// TwinCAT 3 PLC project TcProjectBase
// Title: ATI_KOSTAL_AF2024_AUDI2026_TcProjectBase
// Company: ATI
// Author: Ivana Mishevska
// ProjectVersion: 1.1.0.2
// Description: New library for Festo CMT Drive
// ProgramVersion: 3.1.4024.0
// libraries:
//   KOSTAL.AF2024.Core.FileLogger, * (KOSTAL GmbH & Co.KG)
//   KOSTAL.AF2024.Core.GetSystemTime, * (KOSTAL GmbH & Co.KG)
//   KOSTAL.AF2024.Core.MainControl, * (KOSTAL GmbH & Co.KG)
//   KOSTAL.AF2024.Core.Process, * (KOSTAL GmbH & Co.KG)
//   KOSTAL.AF2024.Core.Settings, * (KOSTAL GmbH & Co.KG)
//   KOSTAL.AF2024.Core.Station, * (KOSTAL GmbH & Co.KG)
//   KOSTAL.AF2024.Core.StringTools, * (KOSTAL GmbH & Co.KG)
//   KOSTAL.AF2024.Core.Text, * (KOSTAL GmbH & Co.KG)
//   KOSTAL.AF2024.Drivers.Actuation.Axis.Festo.CMMT_AS, * (KOSTAL GmbH & Co.KG)
//   KOSTAL.AF2024.Drivers.Actuation.Cylinder, * (KOSTAL GmbH & Co.KG)
//   KOSTAL.AF2024.Drivers.Camera.Cognex_InSight, * (KOSTAL GmbH & Co.KG)
//   KOSTAL.AF2024.Drivers.Camera.I_Camera, * (KOSTAL GmbH & Co.KG)
//   KOSTAL.AF2024.Drivers.Camera.Keyence_IV, * (KOSTAL GmbH & Co.KG)
//   KOSTAL.AF2024.Drivers.Scanner.Cognex.DM260, * (KOSTAL GmbH & Co.KG)
//   KOSTAL.AF2024.Drivers.Scanner.IScanner, * (KOSTAL GmbH & Co.KG)
//   KOSTAL.AF2024.Drivers.Scanner.Keyence_SR, * (KOSTAL GmbH & Co.KG)
//   KOSTAL.AF2024.HMI.I_Hmi, * (KOSTAL GmbH & Co.KG)
//   KOSTAL.AF2024.HMI.WinHMI, * (KOSTAL GmbH & Co.KG)
//   KOSTAL.AF2024.Misc.Counter, * (KOSTAL GmbH & Co.KG)
//   KOSTAL.AF2024.Templates.TextMaster, * (KOSTAL GmbH & Co.KG)
//   KOSTAL.TC3.Device.Axis.FESTO.CMMT_AS.ETC, * (KOSTAL GmbH & Co.KG)
//   Tc2_Standard, * (Beckhoff Automation GmbH)
//   Tc2_System, * (Beckhoff Automation GmbH)
//   Tc2_TcpIp, * (Beckhoff Automation GmbH)
//   Tc2_Utilities, * (Beckhoff Automation GmbH)
//   Tc3_Module, * (Beckhoff Automation GmbH)
//   TcCamera, * (TcNexa)
//   TcCameraKeyenceIX, * (TcNexa)
//   TcProcess, * (TcNexa)
// project tree:
//   00_MainControl_Cell/ FB_MainControlCell.TcPOU, T_E_text_MainControl.TcPOU
//   01_Interface/ I_CustomStationInterface.TcIO
//   02_ControlledStations/ FB_StationBase.TcPOU, FB_StationBaseWithAutomaticSlider.TcPOU, FB_StationBaseWithSlider.TcPOU
//   03_FreeStations/01_Safety/DUTs/ T_E_text_Safety.TcPOU
//   03_FreeStations/01_Safety/ FB_Safety_ST80.TcPOU, FB_SafetyBase.TcPOU, FB_Safety_STAudi.TcPOU, FB_Safety_ST50.TcPOU
//   03_FreeStations/01_Safety/ITFs/ I_Safety.TcIO
//   03_FreeStations/02_Parameters/DUTs/ E_Parameters.TcDUT
//   03_FreeStations/02_Parameters/ FB_ParameterHandler.TcPOU
//   03_FreeStations/02_Parameters/ITFs/ I_Parameters_MainControl.TcIO
//   03_FreeStations/03_TextMaster/DUTs/ T_E_text_Common.TcPOU
//   03_FreeStations/03_TextMaster/ FB_TextMaster.TcPOU
//   03_FreeStations/04_EtherCAT Monitoring/DUTs/ T_E_text_EtherCAT.TcPOU
//   03_FreeStations/04_EtherCAT Monitoring/ FB_EtherCAT_Base.TcPOU
//   03_FreeStations/04_EtherCAT Monitoring/ITFs/ I_EtherCAT.TcIO
//   03_FreeStations/05_Fuse Monitorning/DUTs/ T_E_text_Fuse.TcPOU
//   03_FreeStations/05_Fuse Monitorning/ FB_FuseMonitoringBase.TcPOU
//   03_FreeStations/05_Fuse Monitorning/ITFs/ I_Fuse.TcIO
//   04_ComponentSource/ FB_CounterHandler.TcPOU
//   / GVL_Base_FilesAndFolders.TcGVL, MAIN.TcPOU
//   Version/ Global_Version.TcGVL
// real-time tasks:
//   TASK PlcTask: cycle T#10ms, priority 20, ADS port 350
//   TASK PlcTask1: cycle T#10ms, priority 21, ADS port 351

// ---- 03_FreeStations/02_Parameters/DUTs/E_Parameters.TcDUT
{attribute 'qualified_only'}
{attribute 'strict'}
TYPE E_Parameters :
(
	isLoggerEnabled 				:= 1,
	cylinderTimeout					:= 2,
//	airPressureMin					:= 3,
//	airPressureMax					:= 4,
	numberOfRetries					:= 5
	
);
END_TYPE

// ---- GVL_Base_FilesAndFolders.TcGVL
{attribute 'qualified_only'}
VAR_GLOBAL CONSTANT
	PATH_TEXT_MAIN_CONTROL		: KOSTAL_AF2024_Core_Settings.T_MaxString_UTF8:= 'D:\PLC\Text\MainControl\';
	PATH_TEXT_SAFETY			: KOSTAL_AF2024_Core_Settings.T_MaxString_UTF8:= 'D:\PLC\Text\Safety\';
	PATH_TEXT_ETHERCAT			: KOSTAL_AF2024_Core_Settings.T_MaxString_UTF8:= 'D:\PLC\Text\EtherCAT\';
	PATH_TEXT_FUSE				: KOSTAL_AF2024_Core_Settings.T_MaxString_UTF8:= 'D:\PLC\Text\FuseMonitoring\';
	PATH_PARAMETER_VALUES		: KOSTAL_AF2024_Core_Settings.T_MaxString_UTF8:= 'D:\PLC\Data\parameterValues.json';
	PATH_TEXT_COMMON			: KOSTAL_AF2024_Core_Settings.T_MaxString_UTF8:= 'D:\PLC\Text\Common\';
	PATH_TEXT_MASTER			: KOSTAL_AF2024_Core_Settings.T_MaxString_UTF8:= 'D:\PLC\Text\TextMaster\';
	PATH_TEXT_ARTICLE			: KOSTAL_AF2024_Core_Settings.T_MaxString_UTF8:= 'D:\PLC\Text\Article\';
	PATH_ARTICLES				: KOSTAL_AF2024_Core_Settings.T_MaxString_UTF8:= 'D:\PLC\Article';
	PATH_RESET_COUNTER			: KOSTAL_AF2024_Core_Settings.T_MaxString_UTF8:= 'D:\PLC\Counter\ResettableCounter.json';
	PATH_TOTAL_COUNTER			: KOSTAL_AF2024_Core_Settings.T_MaxString_UTF8:= 'D:\PLC\Counter\TotalCounter.json';
	PATH_LOGGER_PROCESS			: KOSTAL_AF2024_Core_Settings.T_MaxString_UTF8:= 'D:\Log\Process\';
	PATH_LOGGER_SAFETY			: KOSTAL_AF2024_Core_Settings.T_MaxString_UTF8:= 'D:\Log\Safety\';
	PATH_LOGGER_ETHERCAT		: KOSTAL_AF2024_Core_Settings.T_MaxString_UTF8:= 'D:\Log\EtherCAT Diagnostics\';
	PATH_LOGGER_FUSE			: KOSTAL_AF2024_Core_Settings.T_MaxString_UTF8:= 'D:\Log\Fuse Diagnostics\';
	




//	PATH_TEXT_MAIN_CONTROL		: KOSTAL_AF2024_Core_Settings.T_MaxString_UTF8:= 'C:\Users\ATI\Desktop\ST80\PLC\Text\MainControl\';//'D:\PLC\Text\MainControl\';//
//	PATH_TEXT_SAFETY			: KOSTAL_AF2024_Core_Settings.T_MaxString_UTF8:= 'C:\Users\ATI\Desktop\ST80\PLC\Text\Safety\';//'D:\PLC\Text\Safety\';//'
//	PATH_TEXT_ETHERCAT			: KOSTAL_AF2024_Core_Settings.T_MaxString_UTF8:= 'C:\Users\ATI\Desktop\ST80\PLC\Text\EtherCAT\';//'D:\PLC\Text\EtherCAT\';//
//	PATH_TEXT_FUSE				: KOSTAL_AF2024_Core_Settings.T_MaxString_UTF8:= 'C:\Users\ATI\Desktop\ST80\PLC\Text\FuseMonitoring\';//'D:\PLC\Text\FuseMonitoring\';//
//	PATH_PARAMETER_VALUES		: KOSTAL_AF2024_Core_Settings.T_MaxString_UTF8:= 'C:\Users\ATI\Desktop\ST80\PLC\Data\parameterValues.json';//'D:\PLC\Data\parameterValues.json';//
//	PATH_TEXT_COMMON			: KOSTAL_AF2024_Core_Settings.T_MaxString_UTF8:= 'C:\Users\ATI\Desktop\ST80\PLC\Text\Common\';//'D:\PLC\Text\Common\';//
//	PATH_TEXT_MASTER			: KOSTAL_AF2024_Core_Settings.T_MaxString_UTF8:= 'C:\Users\ATI\Desktop\ST80\PLC\Text\TextMaster\';//'D:\PLC\Text\TextMaster\';//
//	PATH_TEXT_ARTICLE			: KOSTAL_AF2024_Core_Settings.T_MaxString_UTF8:= 'C:\Users\ATI\Desktop\ST80\PLC\Text\Article\';//'D:\PLC\Text\Article\';//
//	PATH_ARTICLES				: KOSTAL_AF2024_Core_Settings.T_MaxString_UTF8:= 'C:\Users\ATI\Desktop\ST80\PLC\Article';//'D:\PLC\Article';//
//	PATH_RESET_COUNTER			: KOSTAL_AF2024_Core_Settings.T_MaxString_UTF8:= 'C:\Users\ATI\Desktop\ST80\PLC\Counter\ResettableCounter.json';//
//	PATH_TOTAL_COUNTER			: KOSTAL_AF2024_Core_Settings.T_MaxString_UTF8:= 'D:\PLC\Counter\TotalCounter.json';//'C:\Users\ATI\Desktop\ST80\PLC\Counter\TotalCounter.json';//'D:\PLC\Counter\ResettableCounter.json';//
//	PATH_LOGGER_PROCESS			: KOSTAL_AF2024_Core_Settings.T_MaxString_UTF8:= 'C:\Users\ATI\Desktop\ST80\Log\Process\';//'D:\Log\Process\';//
//	PATH_LOGGER_SAFETY			: KOSTAL_AF2024_Core_Settings.T_MaxString_UTF8:= 'C:\Users\ATI\Desktop\ST80\Log\Safety\';//'D:\Log\Safety\';//
//	PATH_LOGGER_ETHERCAT		: KOSTAL_AF2024_Core_Settings.T_MaxString_UTF8:= 'C:\Users\ATI\Desktop\ST80\Log\EtherCAT Diagnostics\';//'D:\Log\EtherCAT Diagnostics\';//
//	PATH_LOGGER_FUSE			: KOSTAL_AF2024_Core_Settings.T_MaxString_UTF8:= 'C:\Users\ATI\Desktop\ST80\Log\Fuse Diagnostics\';//'D:\Log\Fuse Diagnostics\';//
	
END_VAR

// ---- Version/Global_Version.TcGVL
{attribute 'TcGenerated'}
{attribute 'no-analysis'}
{attribute 'linkalways'}
// This function has been automatically generated from the project information.
VAR_GLOBAL CONSTANT
	{attribute 'const_non_replaced'}
	stLibVersion_ATI_KOSTAL_AF2024_AUDI2026_TcProjectBase : ST_LibVersion := (iMajor := 1, iMinor := 1, iBuild := 0, iRevision := 2, nFlags := 0, sVersion := '1.1.0.2');
END_VAR

// ---- 01_Interface/I_CustomStationInterface.TcIO
INTERFACE I_CustomStationInterface

PROPERTY pressedAbortButton  : BOOL
GET
END_GET
END_PROPERTY

END_INTERFACE

// ---- 03_FreeStations/01_Safety/ITFs/I_Safety.TcIO
INTERFACE I_Safety

PROPERTY PUBLIC doorLock : BOOL
GET
END_GET
SET
END_SET
END_PROPERTY

PROPERTY inHold : BOOL
GET
END_GET
END_PROPERTY

PROPERTY isDoorSafe : BOOL
GET
END_GET
END_PROPERTY

PROPERTY isDoorUsed : BOOL
GET
END_GET
END_PROPERTY

PROPERTY isSafe : BOOL
GET
END_GET
END_PROPERTY

END_INTERFACE

// ---- 03_FreeStations/02_Parameters/ITFs/I_Parameters_MainControl.TcIO
INTERFACE I_Parameters_MainControl

PROPERTY cylinderSensorTimeout : TIME
GET
END_GET
END_PROPERTY

PROPERTY isLoggerEnabled : BOOL
GET
END_GET
END_PROPERTY

PROPERTY numberOfRetries : INT
GET
END_GET
END_PROPERTY

END_INTERFACE

// ---- 03_FreeStations/04_EtherCAT Monitoring/ITFs/I_EtherCAT.TcIO
INTERFACE I_EtherCAT

PROPERTY inError : BOOL
GET
END_GET
END_PROPERTY

END_INTERFACE

// ---- 03_FreeStations/05_Fuse Monitorning/ITFs/I_Fuse.TcIO
INTERFACE I_Fuse

PROPERTY inError : BOOL
GET
END_GET
END_PROPERTY

END_INTERFACE

// ---- 00_MainControl_Cell/FB_MainControlCell.TcPOU
FUNCTION_BLOCK FB_MainControlCell EXTENDS KOSTAL_AF2024_Core_MainControl.FB_MainControl IMPLEMENTS I_CustomStationInterface 
VAR
(*------------------------------------------------------------------------------------------*)
	(* General *)
	_textPath						: KOSTAL_AF2024_Core_Settings.T_MaxString_UTF8;
	_Text							: KOSTAL_AF2024_Core_Text.FB_Handler_Slave;
	_E_Text							: T_E_text_MainControl;
	_setLogRequest					: BOOL;
	_addressHome					: INT;
	_stepDescription				: WSTRING;
	_articleAutoSelection			: BOOL;
	_timerStationsInHome			: Tc2_Standard.TON;
	_tempText						: WSTRING;
	_onAbortButton					: Tc2_Standard.R_TRIG;
//	_pressedAbortButton				: BOOL; 
(*------------------------------------------------------------------------------------------*)
	(* Interface *)
	_IetherCAT						: I_EtherCAT;
	_IfuseMonitroing				: I_Fuse;
	_ISafety						: I_Safety; 
(*------------------------------------------------------------------------------------------*)	 
	(* Hmi *)
	_Hmi							: KOSTAL_AF2024_HMI_WinHMI.FB_MainControl;
	_Hmi_station					: KOSTAL_AF2024_HMI_WinHMI.FB_Page_Station;
(*------------------------------------------------------------------------------------------*)
	(* Mode *)
	_Message						: KOSTAL_AF2024_Core_Process.T_messageText_3_lines;
	_modeAutomaticRequest			: BOOL:= TRUE;
	_modeManualRequest				: BOOL;
	_dataModeRequest				: BOOL;
(*------------------------------------------------------------------------------------------*)
	(* Links *)
	_Ilogger						: KOSTAL_AF2024_Core_FileLogger.I_Logger;
	_Iparameters					: I_Parameters_MainControl;
(*------------------------------------------------------------------------------------------*)
	(* Inputs *)
//	DI_KeySwitch					AT %I* : BOOL;
	DI_KeySwitchAutomatic			AT %I* : BOOL; //2 
	DI_KeySwitchManual				AT %I* : BOOL; //1 
	DI_CheckPressure_PT1			AT %I* : BOOL;
	DI_AbortButton				 	AT %I* : BOOL;
	(* Outputs *)
	DO_AirSupplyOn					AT %Q* : BOOL;
	DO_ReleMainValve_V1				AT %Q* : BOOL;
	DO_ReleMainValve_V2				AT %Q* : BOOL;
	(* Andon Light *)
	DO_AndonLightGreenLamp			AT %Q* : BOOL;
	DO_AndonLightYellowLamp			AT %Q* : BOOL;
	DO_AndonLightRedLamp			AT %Q* : BOOL;
(*------------------------------------------------------------------------------------------*)
END_VAR

VAR CONSTANT
	_STEP_OFF	: INT:= 0;
END_VAR

METHOD PROTECTED _a0_PowerOff
VAR
	_Participant : KOSTAL_AF2024_Core_Settings.T_MaxString;
END_VAR
IF _Step.toggle THEN
	_Message.clear();
	_Hmi.clear();
	_demand.SetUnique_PowerOff();
//	DO_AirSupplyOn:= FALSE;
	DO_ReleMainValve_V1:= FALSE;
	DO_ReleMainValve_V2:= FALSE;
	_setLogRequest:= TRUE;
	_stepDescription:= "PowerOff";
END_IF

// Log
IF _setLogRequest AND _isLogReady() AND _Text.State.ready AND (_Text.LoadedLanguage <> '') THEN
	IF _Log("===START===") THEN 
		_Log(_Text.GetText(Number:= _E_text.off));	
		_setLogRequest:= FALSE;	
	END_IF
END_IF

// Hmi
_Hmi.Button_OnOff.Visible:= FALSE;

IF NOT _Text.State.ready THEN
	_updateHmiText(
		userMessage		:= _Text.GetText(Number:= _E_Text.textHandlerIsNotReady),
		userAction		:= _Text.State.description,
		isErrorMessage	:= FALSE);
ELSIF NOT _Isafety.isSafe THEN
	_updateHmiText(
		userMessage		:= _Text.GetText(Number:= _E_Text.safetyInError),
		userAction		:= "",
		isErrorMessage	:= FALSE);
ELSIF NOT _all_PowerOff(_Participant) THEN
	_updateHmiText(
		userMessage		:= _Text.GetText(Number:= _E_Text.waitForAllOff),
		userAction		:= _Participant,
		isErrorMessage	:= FALSE);
//ELSIF _isAirPressureOk() THEN
//	_Text.ClearVars();
//	_Text.AddVar(Text:= "-1AZ1");
//	_Text.AddVar(Text:= _Text.GetText(Number:= _E_Text.active));
//	_updateHmiText(
//		userMessage		:= _Text.GetText(Number:= _E_Text.systemAirPressure_0_is_1),
//		userAction		:= "",
//		isErrorMessage	:= FALSE);
ELSIF NOT _mode.manual THEN
	_updateHmiText(
		userMessage		:= _Text.GetText(Number:= _E_Text.setManualMode),
		userAction		:= "",
		isErrorMessage	:= FALSE);
ELSE
	_Hmi.Button_OnOff.Visible:= _mode.manual AND NOT _condition.isError();
	
	_Text.ClearVars();
	_Text.AddVar(Text:= _Hmi.Button_OnOff.Text);
	_updateHmiText(
		userMessage		:= _Text.GetText(Number:= _E_Text.onWith_0),
		userAction		:= "",
		isErrorMessage	:= FALSE);

	IF _modeManualRequest AND _Hmi.Button_OnOff.Pulse AND NOT _condition.isError() THEN
		_Step.INC();
	END_IF
END_IF
END_METHOD

METHOD PROTECTED _a1_PowerOn
VAR
	_Participant : KOSTAL_AF2024_Core_Settings.T_MaxString;
END_VAR
IF _step.toggle THEN
	_Hmi.clear();
	_Message.clear();
	_demand.SetUnique_PowerOn();
//	DO_AirSupplyOn:= TRUE;
	DO_ReleMainValve_V1:= TRUE;
	DO_ReleMainValve_V2:= TRUE;
	_log(Text:= _Text.GetText(Number:= _E_Text.powerOn));
	_stepDescription:= "PowerOn";
END_IF

_Hmi.Button_OnOff.Text:= _Text.GetText(Number:= _E_Text.waitForPowerOn);
_Hmi.Button_OnOff.Visible:= TRUE;

//IF NOT _isAirPressureOk() THEN
//	_Text.ClearVars();
////	_Text.AddVar(Text:= INT_TO_WSTRING(_Iparameters.airPressureMin));
////	_Text.AddVar(Text:= INT_TO_WSTRING(AI_AirPressure));
////	_Text.AddVar(Text:= INT_TO_WSTRING(_Iparameters.airPressureMax));
//	_updateHmiText(
//		userMessage		:= _Text.GetText(Number:= _E_Text.waitForAirPressure_0_1_2),
//		userAction		:= "",
//		isErrorMessage	:= FALSE);
IF NOT DI_CheckPressure_PT1 THEN 
	_updateHmiText(
		userMessage		:= "Check pressure",//_Text.GetText(Number:= _E_Text.waitForAirPressure_0_1_2),
		userAction		:= "PT1",
		isErrorMessage	:= FALSE);
ELSIF NOT _all_PowerOn(_Participant) THEN
	_updateHmiText(
		userMessage		:= _Text.GetText(Number:= _E_Text.waitForAllOn),
		userAction		:= _Participant,
		isErrorMessage	:= FALSE);
ELSIF NOT _mode.automatic THEN
	_updateHmiText(
		userMessage		:= _Text.GetText(Number:= _E_Text.setAutomaticMode),
		userAction		:= "",
		isErrorMessage	:= FALSE);
ELSE
	_step.INC();
END_IF
END_METHOD

METHOD PROTECTED _a2_OnToHome
VAR
	_Participant : KOSTAL_AF2024_Core_Settings.T_MaxString;
END_VAR
IF _step.toggle THEN
	_Hmi.clear();
	_demand.SetUnique_OnToHome();
	_log(Text:= _Text.GetText(Number:= _E_Text.onToHomeReleased));
	_stepDescription:= "OnToHome";
END_IF

_Hmi.Button_OnOff.Text:= _Text.GetText(Number:= _E_Text.off);
_Hmi.Button_OnOff.Visible:= TRUE;

IF NOT _all_Home(_Participant) THEN
	_updateHmiText(
		userMessage		:= _Text.GetText(Number:= _E_Text.waitFromHome),
		userAction		:= _Participant,
		isErrorMessage	:= FALSE);
ELSE
	_step.INC();
END_IF
END_METHOD

METHOD PROTECTED _a3_Home
VAR
	_Participant: KOSTAL_AF2024_Core_Settings.T_MaxString;
END_VAR
IF _step.toggle THEN
	_addressHome:= _step.actual;
	_Message.clear();
	_Hmi.clear();
	_demand.SetUnique_Home();
	_log(Text:= _Text.GetText(Number:= _E_Text.stop));
	_stepDescription:= "Home";
END_IF

_Hmi.Button_OnOff.Text:= _Text.GetText(Number:= _E_Text.off);
_Hmi.Button_OnOff.Visible:= TRUE;
_Hmi.Button_RunStop.Text:= _Text.GetText(Number:= _E_Text.start);
_Hmi.Button_RunStop.Visible:= FALSE;

IF NOT _all_Home(_Participant) THEN
	_updateHmiText(
		userMessage		:= _Text.GetText(Number:= _E_Text.participantNotReady),
		userAction		:= _Participant,
		isErrorMessage	:= FALSE);
ELSIF _Hmi.Button_RunStop.Pulse OR NOT _enableStopMode THEN
	_Hmi.Button_RunStop.Visible:= FALSE;
	_step.INC();
ELSE
	_Hmi.Button_RunStop.Visible:= TRUE;
	_updateHmiText(
		userMessage		:= _Text.GetText(Number:= _E_Text.stop),
		userAction		:= _Text.GetText(Number:= _E_Text.readyToStart),
		isErrorMessage	:= FALSE);
END_IF
END_METHOD

METHOD PROTECTED _a4_Run
VAR_INPUT
END_VAR
IF _step.toggle THEN
	_Hmi.clear();
	_demand.SetUnique_Run();
	_log(Text:= _Text.GetText(Number:= _E_Text.busy));
	_stepDescription:= "Run";
END_IF

_Hmi.Button_OnOff.Text:= _Text.GetText(Number:= _E_Text.off);
_Hmi.Button_OnOff.Visible:= TRUE;
_Hmi.Button_RunStop.Text:= _Text.GetText(Number:= _E_Text.stop);
_Hmi.Button_RunStop.Visible:= _enableStopMode;

IF _Hmi.Button_RunStop.Pulse AND _enableStopMode THEN
	_step.INC();
//ELSIF NOT _isAirPressureOk() THEN
//	_updateHmiText(
//		userMessage		:= "Air pressure out of limits",
//		userAction		:= "",
//		isErrorMessage	:= TRUE);
//	_step.init();	
//ELSIF (_IetherCAT <> 0) AND_THEN _IetherCAT.inError THEN
//	_updateHmiText(
//		userMessage		:= "EtherCAT in fault",
//		userAction		:= "",
//		isErrorMessage	:= TRUE);
//	_step.init();	
//ELSIF (_IfuseMonitroing <> 0) AND_THEN _IfuseMonitroing.inError THEN
//	_updateHmiText(
//		userMessage		:= "Fuse in fault",
//		userAction		:= "",
//		isErrorMessage	:= TRUE);
//	_step.init();	
ELSE
	_tempText:= "";
//	IF (_IArticle <> 0) THEN
//		IF _IArticle.LoadedArticle.isVariantTypeGen6x THEN
//			_tempText:= "Selected article: Gen6x";
//		ELSIF _IArticle.LoadedArticle.isProductTypeGen6 THEN
//			_tempText:= "Selected article: Gen6";
//		ELSIF _IArticle.LoadedArticle.isProductTypeGen7 THEN
//			_tempText:= "Selected article: Gen7";
//		ELSIF _IArticle.LoadedArticle.isProductTypeVan THEN
//			_tempText:= "Selected article: Van";
//		END_IF
//	END_IF

	_updateHmiText(
		userMessage		:= _Text.GetText(Number:= _E_Text.run),
		userAction		:= _tempText,
		isErrorMessage	:= FALSE);
END_IF
END_METHOD

METHOD PROTECTED _a5_RunToHome
VAR
	_Participant: KOSTAL_AF2024_Core_Settings.T_MaxString;
END_VAR
IF _step.toggle THEN
	_Message.clear();
	_Hmi.clear();
	_demand.SetUnique_RunToHome();
	_log(Text:= _Text.GetText(Number:= _E_Text.lastCycle));
	_stepDescription:= "RunToHome";
END_IF

_Hmi.Button_OnOff.Text:= _Text.GetText(Number:= _E_Text.off);
_Hmi.Button_OnOff.Visible:= TRUE;
_Hmi.Button_RunStop.Text:= _Text.GetText(Number:= _E_Text.start);
_Hmi.Button_RunStop.Visible:= TRUE;

IF _Hmi.Button_RunStop.Pulse OR NOT _enableStopMode THEN
	_step.DEC();
ELSIF _all_Home(_Participant) THEN
	_step.set(request:= _addressHome);
ELSE
	_updateHmiText(
		userMessage		:= _Text.GetText(Number:= _E_Text.participantNotReady),
		userAction		:= _Participant,
		isErrorMessage	:= FALSE);
END_IF
END_METHOD

METHOD PROTECTED _aX_Fail
VAR_INPUT
END_VAR
_demand.clear();

_Message.clear();
_Text.ClearVars();
_Text.AddVar(Text:= INT_TO_WSTRING(_Step.actual));
_Message.line_01:= _Text.GetText(Number:= _E_Text.step_0_doesNotExist);
_condition.setMessage(
	priority:= _condition.PriorityLevel_Error + 1000,
	message:= _Message);
	
IF _Step.toggle THEN
	_Log(Text:= _Message.toString());
END_IF

_Step.init();
END_METHOD

METHOD PROTECTED _checkIfSamePosition : BOOL
VAR_INPUT
	actualPosition 			: LREAL;
	targetPosotion			: LREAL;
END_VAR
IF (actualPosition >= (targetPosotion - 1)) AND (actualPosition <= (targetPosotion + 1)) THEN 
	_checkIfSamePosition:= TRUE;
ELSE 
	_checkIfSamePosition:= FALSE;
END_IF
END_METHOD

METHOD PROTECTED _getIdAsString : KOSTAL_AF2024_Core_Settings.T_MaxString
VAR
	_temp 		: KOSTAL_AF2024_Core_StringTools.FB_Concat;
END_VAR
_temp.Clear();
_temp.addContent(Text:= _ID.name);
_temp.addContent(Text:= "(");
_temp.addContent(Text:= DINT_TO_WSTRING(_ID.key));
_temp.addContent(Text:= ")");
_getIdAsString:= _temp.getResult();
_temp.Clear();
END_METHOD

METHOD PROTECTED _globalError
VAR_INPUT
END_VAR
END_METHOD

METHOD PROTECTED _handleAndonLight
VAR
	_Participant	: KOSTAL_AF2024_Core_Settings.T_MaxString;
END_VAR
IF NOT _Isafety.isSafe THEN
	_timerStationsInHome(IN:= FALSE);
	DO_AndonLightGreenLamp:= FALSE;
	DO_AndonLightYellowLamp:= FALSE;
	DO_AndonLightRedLamp:= TRUE;
ELSIF _mode.manual THEN
	_timerStationsInHome(IN:= FALSE);
	DO_AndonLightGreenLamp:= FALSE;
	DO_AndonLightYellowLamp:= TRUE;
	DO_AndonLightRedLamp:= FALSE;
ELSIF _all_Home(_Participant) THEN
	_timerStationsInHome(IN:= TRUE, PT:= T#1S);
	DO_AndonLightYellowLamp:= FALSE;
	DO_AndonLightRedLamp:= FALSE;
	IF _timerStationsInHome.Q THEN
		_timerStationsInHome(IN:= FALSE);
		DO_AndonLightGreenLamp:= NOT DO_AndonLightGreenLamp;
	END_IF
ELSE
	_timerStationsInHome(IN:= FALSE);
	DO_AndonLightGreenLamp:= TRUE;
	DO_AndonLightYellowLamp:= FALSE;
	DO_AndonLightRedLamp:= FALSE;
END_IF
END_METHOD

METHOD PROTECTED _hmiDefine
VAR
	_Participant: KOSTAL_AF2024_Core_Settings.T_MaxString;
END_VAR
_Hmi.FBmain();
_Hmi_station.FBmain();

// General
_Hmi.Name:= "";
_Hmi.linkMainControl(THIS^);

_Hmi_station.Name:= Tc2_Standard.WCONCAT(
	STR1:= _Text.GetText(Number:= _E_Text.name),
	STR2:= " [");
_Hmi_station.Name:= Tc2_Standard.WCONCAT(
	STR1:= _Hmi_station.Name,
	STR2:= STRING_TO_WSTRING(stLibVersion_ATI_KOSTAL_AF2024_AUDI2026_TcProjectBase.sVersion));
_Hmi_station.Name:= Tc2_Standard.WCONCAT(
	STR1:= _Hmi_station.Name,
	STR2:= "]");

// Mode handling
_mode.manual:= _modeManualRequest;
_mode.automatic:= _modeAutomaticRequest AND NOT _Isafety.inHold;

// Buttons 
_Hmi.Button_Parameters.Visible:= (NOT DI_KeySwitchAutomatic AND NOT DI_KeySwitchManual) AND _dataModeRequest;//_mode.automatic
_Hmi.Button_Article.Visible:= _mode.manual AND _demand.Run; //AND (_Hmi.UserLevel >= KOSTAL_AF2024_HMI_I_Hmi.E_UserLevel.service);
_Hmi.Button_RunStop.Visible:= _enableStopMode;
_Hmi.ManualDeviceControl:= _mode.manual AND _demand.Run AND (_Hmi.UserLevel >= KOSTAL_AF2024_HMI_I_Hmi.E_UserLevel.service);


_Hmi.Button_Door.Visible:= _ISafety.isDoorUsed;
IF _Hmi.Button_Door.Pulse THEN
	_ISafety.doorLock:= NOT _ISafety.doorLock;
END_IF
_Hmi.statusDoor_safe:= _ISafety.isDoorSafe;

_Hmi_station.Button_Escape.Visible:= _condition.isError() AND _modeManualRequest;
_Hmi_station.Button_Escape.Text:= _Text.GetText(Number:= _E_Text.reset);

// Message
_Hmi_station.Text.line_01:= _condition.Message.line_01;
_Hmi_station.Text.line_02:= _condition.Message.line_02;
_Hmi_station.Text.line_03:= _condition.Message.line_03;
_Hmi_station.Status.CopyFrom(IN:= _condition);
END_METHOD

METHOD PROTECTED _isLogReady  : BOOL
VAR_INPUT
END_VAR
IF (_Ilogger = 0) THEN RETURN; END_IF
_isLogReady:= _Ilogger.State.success;
END_METHOD

METHOD PROTECTED _log : BOOL
VAR_INPUT
	Text			  : KOSTAL_AF2024_Core_Settings.T_MaxString;
END_VAR
IF (Text = "") THEN RETURN; END_IF
IF (_Iparameters <> 0) AND_THEN NOT _Iparameters.isLoggerEnabled THEN RETURN; END_IF
IF (_Ilogger = 0) THEN RETURN; END_IF
IF NOT _Ilogger.State.success THEN RETURN; END_IF

_Ilogger.ID:= _getIdAsString();
_Ilogger.name:= _Text.GetText(Number:= _E_Text.name);
_Ilogger.stepNumber:= _Step.actual;

_log:= _Ilogger.addLine(line:= Text);
END_METHOD

METHOD _modeHandler
VAR_INPUT
END_VAR
_mode.automatic:= (_modeAutomaticRequest OR DI_KeySwitchAutomatic) AND NOT _condition.isError() AND NOT _Isafety.inHold AND NOT _dataModeRequest; 
_mode.manual:= _modeManualRequest AND NOT _dataModeRequest;
END_METHOD

METHOD PROTECTED _modeRequest
VAR_INPUT
END_VAR
_Hmi.Button_Auto.Visible:= TRUE;
_Hmi.Button_Manual.Visible:= TRUE;
IF _Hmi.Button_Auto.Pulse OR DI_KeySwitchAutomatic THEN	
	_modeAutomaticRequest:= TRUE;	
	_modeManualRequest:= FALSE;
	_dataModeRequest:= FALSE;
ELSIF _Hmi.Button_Manual.Pulse OR DI_KeySwitchManual THEN	
	_modeAutomaticRequest:= FALSE;	
	_modeManualRequest:= TRUE;
	_dataModeRequest:= FALSE;
ELSIF NOT DI_KeySwitchAutomatic AND NOT DI_KeySwitchManual THEN 
//	_Hmi.Button_Auto.Visible:= TRUE;
//	_Hmi.Button_Manual.Visible:= TRUE;
	_dataModeRequest:= TRUE;
	_modeAutomaticRequest:= FALSE;
	_modeManualRequest:= FALSE;
END_IF
END_METHOD

METHOD PROTECTED _parameterControl : BOOL
VAR_INPUT
END_VAR
_parameterControl:= TRUE;
END_METHOD

METHOD PROTECTED _resetCondition  
VAR_INPUT
END_VAR
IF _condition.isError() THEN
	IF _Hmi_station.Button_Escape.Pulse THEN
		_condition.clear();
	END_IF
ELSE
	_condition.clear();
END_IF
END_METHOD

METHOD PROTECTED _stepHeader
VAR_INPUT
END_VAR
//Switch off in case of off command or safety error
IF _step.actual > _STEP_OFF THEN
	IF _hmi.Button_OnOff.Pulse THEN	
		_step.init();
	ELSIF NOT _Isafety.IsSafe THEN
		_step.init();
	END_IF
END_IF
//Call Step sequence header
_step.Header();
END_METHOD

METHOD PROTECTED _steps
VAR_INPUT
END_VAR
_stepHeader();

CASE _Step.actual OF
	0:	_a0_PowerOff();
	1:	_a1_PowerOn();
	2:	_a2_OnToHome();
	3:	_a3_Home();
	4:	_a4_Run();
	5:	_a5_RunToHome();
ELSE
	_aX_Fail();
END_CASE
END_METHOD

METHOD PROTECTED _textReader : BOOL
VAR_INPUT
END_VAR
_Text.Path:= _textPath;
_Text.FBmain();

IF _Text.State.fail THEN
	_Message.clear();
	_Message.line_01:= "TextHandler";
	_Message.line_02:= _Text.State.description;
	_condition.setMessage(
		priority:= _condition.PriorityLevel_Error,
		message	:= _Message);
ELSIF NOT _Text.Valid THEN
	_Message.clear();
	_Message.line_01:= "TextHandler";
	_Message.line_02:= _Text.State.description;
	_condition.setMessage(
		priority:= _condition.PriorityLevel_MasterMessage + 999,
		message	:= _Message);
END_IF

IF _Text.LoadedLanguage <> '' THEN
	_textReader:= TRUE;
END_IF
END_METHOD

METHOD PROTECTED _updateHmiText
VAR_INPUT
	userMessage		: WSTRING;
	userAction		: WSTRING;
	isErrorMessage	: BOOL;
END_VAR
_message.clear();

_Text.ClearVars();
_Text.AddVar(Text:= INT_TO_WSTRING(_step.actual));
_Text.AddVar(Text:= _stepDescription);
_Text.AddVar(Text:= "0");
_message.line_01:= _Text.GetText(Number:= _E_Text.step_0_actual_1);
_message.line_02:= userMessage;
_message.line_03:= userAction;
IF isErrorMessage AND NOT _condition.isError() THEN
	_log(Text:= _message.toString());
END_IF

IF isErrorMessage THEN
	_condition.setMessage(
		priority:= _condition.PriorityLevel_Error,
		message	:= _message);
ELSIF (userAction <> "") THEN
	_condition.setMessage(
		priority:= _condition.PriorityLevel_Message,
		message	:= _message);
ELSE
	_condition.setMessage(
		priority:= _condition.PriorityLevel_Text,
		message	:= _message);
END_IF
END_METHOD

PROPERTY articleAutoSelection : BOOL
GET
articleAutoSelection:= _articleAutoSelection;
END_GET
SET
_articleAutoSelection:= articleAutoSelection;
END_SET
END_PROPERTY

METHOD FB_init : BOOL
VAR_INPUT
	bInitRetains 		: BOOL; // if TRUE, the retain variables are initialized (warm start / cold start)
	bInCopyCode 		: BOOL;  // if TRUE, the instance afterwards gets moved into the copy code (online change)
	EnableStopMode		: BOOL;
	CommonText			: KOSTAL_AF2024_Core_Text.I_Text;
	textPath			: KOSTAL_AF2024_Core_Settings.T_MaxString_UTF8;
	Parameters			: I_Parameters_MainControl;
	Safety				: I_Safety;
	EtherCAT			: I_EtherCAT;
	Fuse				: I_Fuse;
	Logger				: KOSTAL_AF2024_Core_FileLogger.I_Logger;
//	Article				: I_Article;
END_VAR
THIS^._enableStopMode:= EnableStopMode;
THIS^._Text.linkCommonText(Common:= CommonText);
THIS^._textPath:= textPath;
THIS^._Iparameters:= Parameters;
THIS^._Isafety:= Safety;
THIS^._IetherCAT:= EtherCAT;
THIS^._IfuseMonitroing:= Fuse;
THIS^._Ilogger:= Logger;
END_METHOD

METHOD PUBLIC FBmain 
VAR_INPUT
END_VAR
_modeRequest();

IF NOT _parameterControl() THEN RETURN; END_IF
_hmiDefine();
_resetCondition();
_handleAndonLight();

IF NOT _TextReader() THEN RETURN; END_IF

_globalError();
_modeHandler();
_steps();

_onAbortButton(CLK:= DI_AbortButton);
END_METHOD

PROPERTY language : KOSTAL_AF2024_HMI_I_Hmi.T_LANGUAGENAME
GET
language:= _Hmi.Language;
END_GET
END_PROPERTY

{warning 'add property implementation'}
PROPERTY pressedAbortButton : BOOL
GET
pressedAbortButton:= _onAbortButton.Q;
END_GET
END_PROPERTY

PROPERTY user : KOSTAL_AF2024_HMI_I_Hmi.E_UserLevel
GET
user:= _Hmi.UserLevel;
END_GET
END_PROPERTY

END_FUNCTION_BLOCK

// ---- 00_MainControl_Cell/T_E_text_MainControl.TcPOU
FUNCTION_BLOCK T_E_text_MainControl EXTENDS KOSTAL_AF2024_Core_Text.T_E_Text
VAR
END_VAR

PROPERTY busy : KOSTAL_AF2024_Core_Text.ST_E_Text
GET
busy.Number:= 36;
END_GET
END_PROPERTY

PROPERTY lastCycle : KOSTAL_AF2024_Core_Text.ST_E_Text
GET
lastCycle.Number:= 37;
END_GET
END_PROPERTY

PROPERTY name : KOSTAL_AF2024_Core_Text.ST_E_Text
GET
name.Number:= 2;
END_GET
END_PROPERTY

PROPERTY nextPage : KOSTAL_AF2024_Core_Text.ST_E_Text
GET
nextPage.Number:= 61;
END_GET
END_PROPERTY

PROPERTY off : KOSTAL_AF2024_Core_Text.ST_E_Text
GET
off.Source:= KOSTAL_AF2024_Core_Text.E_Source.Common;
off.Number:= 2;
END_GET
END_PROPERTY

PROPERTY onToHomeReleased : KOSTAL_AF2024_Core_Text.ST_E_Text
GET
onToHomeReleased.Source:= KOSTAL_AF2024_Core_Text.E_Source.Common;
onToHomeReleased.Number:= 42;
END_GET
END_PROPERTY

PROPERTY onWith_0 : KOSTAL_AF2024_Core_Text.ST_E_Text
GET
onWith_0.Source:= KOSTAL_AF2024_Core_Text.E_Source.Common;
onWith_0.Number:= 65;
END_GET
END_PROPERTY

PROPERTY participantNotReady : KOSTAL_AF2024_Core_Text.ST_E_Text
GET
participantNotReady.Number:= 12;
END_GET
END_PROPERTY

PROPERTY powerOn : KOSTAL_AF2024_Core_Text.ST_E_Text
GET
powerOn.Number:= 44;
END_GET
END_PROPERTY

PROPERTY previousPage : KOSTAL_AF2024_Core_Text.ST_E_Text
GET
previousPage.Number:= 60;
END_GET
END_PROPERTY

PROPERTY readyToStart : KOSTAL_AF2024_Core_Text.ST_E_Text
GET
readyToStart.Number:=35;
END_GET
END_PROPERTY

PROPERTY refresh : KOSTAL_AF2024_Core_Text.ST_E_Text
GET
refresh.Number:= 62;
END_GET
END_PROPERTY

PROPERTY reset : KOSTAL_AF2024_Core_Text.ST_E_Text
GET
reset.Source:= Kostal_AF2024_Core_Text.E_Source.Common;
reset.Number:= 7;
END_GET
END_PROPERTY

PROPERTY run : KOSTAL_AF2024_Core_Text.ST_E_Text
GET
run.Number:= 5;
END_GET
END_PROPERTY

PROPERTY safetyInError : KOSTAL_AF2024_Core_Text.ST_E_Text
GET
safetyInError.Number:= 30;
END_GET
END_PROPERTY

PROPERTY setAutomaticMode : KOSTAL_AF2024_Core_Text.ST_E_Text
GET
setAutomaticMode.Number:=41;
END_GET
END_PROPERTY

PROPERTY setManualMode : KOSTAL_AF2024_Core_Text.ST_E_Text
GET
setManualMode.Number:= 40;
END_GET
END_PROPERTY

PROPERTY start : KOSTAL_AF2024_Core_Text.ST_E_Text
GET
start.Source:= KOSTAL_AF2024_Core_Text.E_Source.Common;
start.Number:= 5;
END_GET
END_PROPERTY

PROPERTY step_0_actual_1 : KOSTAL_AF2024_Core_Text.ST_E_Text
GET
step_0_actual_1.Source:= KOSTAL_AF2024_Core_Text.E_Source.Common;
step_0_actual_1.Number:= 11;
END_GET
END_PROPERTY

PROPERTY step_0_doesNotExist : KOSTAL_AF2024_Core_Text.ST_E_Text
GET
step_0_doesNotExist.Source:= KOSTAL_AF2024_Core_Text.E_Source.Common;
step_0_doesNotExist.Number:= 12;
END_GET
END_PROPERTY

PROPERTY stop : KOSTAL_AF2024_Core_Text.ST_E_Text
GET
stop.Source:= KOSTAL_AF2024_Core_Text.E_Source.Common;
stop.Number:= 4;
END_GET
END_PROPERTY

PROPERTY textHandlerIsNotReady : KOSTAL_AF2024_Core_Text.ST_E_Text
GET
textHandlerIsNotReady.Source:= KOSTAL_AF2024_Core_Text.E_Source.Common;
textHandlerIsNotReady.Number:= 20;
END_GET
END_PROPERTY

PROPERTY waitForAirPressure_0_1_2 : KOSTAL_AF2024_Core_Text.ST_E_Text
GET
waitForAirPressure_0_1_2.Number:= 31;
END_GET
END_PROPERTY

PROPERTY waitForAllOff : KOSTAL_AF2024_Core_Text.ST_E_Text
GET
waitForAllOff.Number:= 10;
END_GET
END_PROPERTY

PROPERTY waitForAllOn : KOSTAL_AF2024_Core_Text.ST_E_Text
GET
waitForAllOn.Number:= 11;
END_GET
END_PROPERTY

PROPERTY waitForPowerOn : KOSTAL_AF2024_Core_Text.ST_E_Text
GET
waitForPowerOn.Number:= 13;
END_GET
END_PROPERTY

PROPERTY waitFromHome : KOSTAL_AF2024_Core_Text.ST_E_Text
GET
waitFromHome.Number:= 43;
END_GET
END_PROPERTY

END_FUNCTION_BLOCK

// ---- 02_ControlledStations/FB_StationBase.TcPOU
FUNCTION_BLOCK ABSTRACT FB_StationBase EXTENDS KOSTAL_AF2024_Core_Station.FB_Station_Controlled 
VAR PERSISTENT
	_isCameraMasterDone					: BOOL;
	_lastCameraMasterTime				: DINT;	
END_VAR                         		
VAR                             		
	(* General *)  	            		
	_Hmi_station						: KOSTAL_AF2024_HMI_WinHMI.FB_Page_Station;
	_E_TextCommon						: T_E_text_Common;
	_IgetTime							: KOSTAL_AF2024_Core_GetSystemTime.I_TimeSource;
	_isDevicesInit						: BOOL;
	_cylinderInManualMode				: BOOL;
	_manualModeInterlock				: BOOL;
	_onPowerOff							: Tc2_Standard.R_TRIG;
	_onNagaraSwitch						: Tc2_Standard.R_TRIG;
//	_onAbortButton						: Tc2_Standard.R_TRIG;
	_timerCycleTimer					: Tc2_Standard.TON;
	_addressRestart						: INT;
	_tempText							: KOSTAL_AF2024_Core_Settings.T_MaxString_UTF8;
	_isHomeControkOk					: BOOL;
	_TextSplitter						: KOSTAL_AF2024_Core_StringTools.FB_Split;
	_cycleTime							: TIME;
	_CloseAllSockets					: Tc2_TcpIp.FB_SocketCloseAll;
	_isTcpIpInit						: BOOL;
	_WritePersistentData				: Tc2_Utilities.WritePersistentData;
	(* Camera master *)         		
	_onShiftChange						: Tc2_Standard.R_TRIG;
	_cameraMasterOnStartupDone			: BOOL;
	_isCameraMasterBadPartDone			: BOOL;
	_isCameraMasterGoodPartDone			: BOOL;
	_timeForMaster						: BOOL; 
	(* Process *)               		
	_isStepInit							: BOOL;
	_onStateHome						: Tc2_Standard.R_TRIG;
	_SubStep							: KOSTAL_AF2024_Core_Process.FB_processStep_Flow;
	_lastSubStep						: INT;
	_stepDescription					: KOSTAL_AF2024_Core_Settings.T_MaxString;
	_subStepError						: KOSTAL_AF2024_Core_Settings.T_MaxString;
	_subStepMessage						: KOSTAL_AF2024_Core_Settings.T_MaxString;
	_onSubStepRetryAbort				: Tc2_Standard.R_TRIG;
	_retryPartsInSeries					: INT;
	_partOk								: BOOL;
	_partNok							: BOOL;
	(* Interface *)             		
	_IresettableCounter					: KOSTAL_AF2024_Misc_Counter.I_T_CounterSet;
	_ItotalCounter						: KOSTAL_AF2024_Misc_Counter.I_T_CounterSet;
	_IparametersBase					: I_Parameters_MainControl;
	_IStation							: I_CustomStationInterface; 
	(* Sensors *)
	DI_NagaraSwitch				 AT %I* : BOOL; 
//	DI_AbortButton				 AT %I* : BOOL;
	(* Process Light *)
	DO_ProcessLightGreenLamp	 AT %Q* : BOOL;
	DO_ProcessLightRedLamp		 AT %Q* : BOOL;
	DO_ProcessLightYellowLamp	 AT %Q* : BOOL;
	DO_ProcessLightBlueLamp		 AT %Q* : BOOL;
	(* IX camera *)
	 _InternalResponse					: TcNexa_Components_TcProcess.FB_MethodResponse;
	(* SPC counter *)
	_counterForSCPmode					: INT;
	_isSPCmodeActive					: BOOL;
END_VAR
VAR CONSTANT
	(* Step *)
	_ADDRESS_POWEROFF					: INT:= 0;
	_ADDRESS_READY						: INT:= 30;	
	_ADDRESS_PASS						: INT:= 100;
	_ADDRESS_FAIL						: INT:= 200;
	_ADDRESS_SPCMODE					: INT:= 300;
	_ADDRESS_RUNOUT						: INT:= 350;
	_ADDRESS_CAMERA_MASTER				: INT:= 400;
	
	(* Sub Step *)              		
	_SUB_ADDRESS_PASS					: INT:= 600;
	_SUB_ADDRESS_RETRY_ABORT			: INT:= 700;
	_SUB_ADDRESS_ABORT					: INT:= 800;
	(* General *)               		
	_UNLIMITED_RETRY_NUMBER				: INT:= -1;
END_VAR

METHOD PROTECTED _a0_Fail
VAR_INPUT
END_VAR
_Text.ClearVars();
_Text.AddVar(Text:= INT_TO_WSTRING(_step.actual));

_message.clear();
_message.line_01:= _Text.GetText(Number:= _E_TextCommon.step_0_DoesNotExist);
_condition.setMessage(
	priority	:= _condition.PriorityLevel_Error + 1000,
	message		:= _message);
_log(Text:= _message.toString());
END_METHOD

METHOD PROTECTED _a1_000_PowerOff
VAR_INPUT
END_VAR
IF _step.toggle THEN
	_Hmi_station.clear();
	_log(Text:= _Text.GetText(Number:= _E_TextCommon.off));
	_state.SetUnique_PowerOff();
	_stepDescription:= "PowerOff";
END_IF

_condition.clear();
_message.clear();
_Hmi_station.clear_controls();

_updateHmiText(
	userMessage		:= _Text.GetText(Number:= _E_TextCommon.off), 
	userAction		:= "", 
	isErrorMessage	:= FALSE);

IF _mainControl.Demand.PowerOn THEN
	_log(Text:= _Text.GetText(Number:= _E_TextCommon.on));
	_step.INC();
ELSIF _Hmi_station.Button_OnOff.Pulse THEN
	;
END_IF
END_METHOD

METHOD PROTECTED _a1_001_PowerOn
VAR_INPUT
END_VAR
IF _step.toggle THEN
	_state.SetUnique_PowerOn();
	_stepDescription:= "PowerOn";
END_IF

_updateHmiText(
	userMessage		:= _Text.GetText(Number:= _E_TextCommon.on), 
	userAction		:= "", 
	isErrorMessage	:= FALSE);

IF _mainControl.Demand.OnToHome THEN
	_step.Condition:= TRUE;
END_IF

_step.Control();
END_METHOD

METHOD PROTECTED _a1_X_Finish
VAR_INPUT
END_VAR
IF _step.toggle THEN
	_state.SetUnique_Finish();
END_IF

_step.set(request:= _ADDRESS_READY);
END_METHOD

METHOD PROTECTED ABSTRACT _a2_002_HomeStation
VAR_INPUT
END_VAR
END_METHOD

METHOD PROTECTED _a2_030_Ready
VAR_INPUT
END_VAR
IF _step.toggle THEN
	_partOk:= FALSE;
	_partNok:= FALSE;
	_state.SetUnique_Home();
	_stepDescription:= "Ready";
END_IF

_isHomeControkOk:= _a2_030_Ready_HomeControl();

(* Machine is in stop state *)
IF NOT _mainControl.Demand.Run THEN
	_Text.ClearVars();
	_Text.AddVar(Text:= _Text.GetText(Number:= _E_TextCommon.stop));
	_updateHmiText(
		userMessage		:= _Text.GetText(Number:= _E_TextCommon.mainControlIsIn_0_state), 
		userAction		:= "", 
		isErrorMessage	:= FALSE);
ELSIF _cylinderInManualMode THEN
	_updateHmiText(
		userMessage		:= _Text.GetText(Number:= _E_TextCommon.stationInManualMode), 
		userAction		:= _Text.GetText(Number:= _E_TextCommon.cylinderInManualMode), 
		isErrorMessage	:= FALSE);
ELSIF _isHomeControkOk THEN
	_a2_030_Ready_ConditionControl();
END_IF

_step.Control();

IF _step.Done THEN
	_state.SetUnique_Busy();
END_IF
END_METHOD

METHOD PROTECTED ABSTRACT _a2_030_Ready_ConditionControl
VAR_INPUT
END_VAR
END_METHOD

METHOD PROTECTED ABSTRACT _a2_030_Ready_HomeControl : BOOL
VAR_INPUT
END_VAR
END_METHOD

METHOD PROTECTED _a2_X_CognexCameraTrigerTCPIP : BOOL
VAR_INPUT
	Camera				 : KOSTAL_AF2024_Drivers_Camera_Cognex_InSight.I_InSight_TcpIp;
	targetProgramNum	 : UINT;
	isCameraEnable		 : BOOL;
	cameraName			 : STRING;
	
END_VAR
IF _step.toggle THEN 
	_stepDescription:= "CognexCameraCheck";
END_IF

(* Check Camera Ready *)
IF _SubStep.isActive(0) THEN 
	_addressRestart:= _SubStep.actual;
	IF NOT isCameraEnable THEN 
		_a2_X_CognexCameraTrigerTCPIP:= TRUE;
//		_SubStep.set(request:= _SUB_ADDRESS_PASS);
	ELSIF NOT Camera.State.ready THEN 
		_updateHmiTextWithCameraNotReady(name:= STRING_TO_WSTRING( cameraName));
	ELSE 
		_addressRestart:= _SubStep.actual;
		_SubStep.INC();
	END_IF
END_IF
(* Camera triger *) //Ima program number i program name 
IF _SubStep.isActive(1) THEN 
	IF NOT Camera.Ex_Trigger_ProgramNumber(ProgramNumber:= targetProgramNum) THEN 
		_updateHmiTextWithCameraBusy(name:= STRING_TO_WSTRING(cameraName));
	ELSIF NOT Camera.State.finish THEN 
		_updateHmiTextWithCameraBusy(name:= STRING_TO_WSTRING(cameraName));
	ELSIF NOT Camera.State.pass THEN 
		_getCameraErrorTexts(
			name		:= STRING_TO_WSTRING( cameraName),
			description	:= Camera.State.description);
		_a2_X_CognexCameraTrigerTCPIP:= FALSE;
//		_SubStep.set(request:= _SUB_ADDRESS_RETRY_ABORT);
	ELSE 
//		_SubStep.set(request:= _SUB_ADDRESS_PASS);
		_a2_X_CognexCameraTrigerTCPIP:= TRUE;
	END_IF
END_IF

(* Pass *)
//IF _SubStep.isActive(_SUB_ADDRESS_PASS) THEN
////	_step.Condition:= TRUE;
//	_SubStep.INC();
//END_IF
(* Fail *)
//IF _SubStep.isActive(_SUB_ADDRESS_RETRY_ABORT) THEN
//	_retryAbort(
//		numOfTargetRetries	:= _IparametersBase.numberOfRetries, 
//		retryAddress		:= _addressRestart, 
//		abortAddress		:= _ADDRESS_RUNOUT);
//END_IF

//_step.Control();
END_METHOD

METHOD PROTECTED _a2_X_CognexReaderScanCode
VAR_INPUT
	Scanner			: KOSTAL_AF2024_Drivers_Scanner_Cognex_DM260.I_Scanner;
	isScanerEnable	: BOOL;
END_VAR
VAR_OUTPUT
	SFC				: KOSTAL_AF2024_Core_Settings.T_MaxString_UTF8;
END_VAR
//Da se proba dali kje raboti vaka ako ne kje treba enable na nekoj setting da se napravi 
//Ili tcp ip 

IF _step.toggle THEN 
	_stepDescription:= "ScanCode";
END_IF

(* Wait until scanner is ready *)
IF _SubStep.isActive(0) THEN 
	_addressRestart:= _SubStep.actual;
	IF NOT isScanerEnable THEN 
		SFC:= '';
		_SubStep.set(request:= _SUB_ADDRESS_PASS);
	ELSIF NOT Scanner.State.ready THEN 
		_Text.ClearVars();
		_text.AddVar("41A1");
		_updateHmiText(
			userMessage		:= _Text.GetText(Number:= _E_TextCommon.scanner_0_failed),
			userAction		:= _Text.GetText(Number:= _E_TextCommon.scanner_0_notReady),
			isErrorMessage	:= FALSE);
	ELSE 
		_SubStep.INC();
	END_IF
END_IF

(* Execute *)
IF _SubStep.isActive(1) THEN 
	IF NOT Scanner.Ex_Scan() THEN 
		_Text.ClearVars();
		_text.AddVar("41A1");
		_updateHmiText(
			userMessage		:= _Text.GetText(Number:= _E_TextCommon.scanner_0_busy),
			userAction		:= "",
			isErrorMessage	:= FALSE);
	ELSIF NOT Scanner.State.finish THEN 
		_Text.ClearVars();
		_text.AddVar("41A1");
		_updateHmiText(
			userMessage		:= _Text.GetText(Number:= _E_TextCommon.scanner_0_busy),
			userAction		:= "",
			isErrorMessage	:= FALSE);
	ELSIF NOT Scanner.State.pass THEN 
		_Text.ClearVars();
		_text.AddVar("41A1");
		_updateHmiText(
			userMessage		:= _Text.GetText(Number:= _E_TextCommon.scanner_0_inError),
			userAction		:= Scanner.State.description,
			isErrorMessage	:= FALSE);
		_SubStep.set(request:= _SUB_ADDRESS_RETRY_ABORT);
	ELSIF (Scanner.CodeGet(1) = '') OR (Scanner.CodeGet(1) = 'ERROR') OR (Scanner.CodeGet(1) = 'NONE') THEN 
		_Text.ClearVars();
		_updateHmiText(
			userMessage		:= _Text.GetText(Number:= _E_TextCommon.scanner_0_failed),
			userAction		:= _Text.GetText(Number:= _E_TextCommon.scanner_0_noCode),
			isErrorMessage	:= FALSE);
		_SubStep.set(request:= _SUB_ADDRESS_RETRY_ABORT);
	ELSE 
		_SubStep.set(request:= _SUB_ADDRESS_PASS);	
	END_IF
END_IF

(* Pass *) 
IF _SubStep.isActive(_SUB_ADDRESS_PASS) THEN 
	SFC:= Scanner.CodeGet(number:= 1);
	_step.Condition:= TRUE;
END_IF
(* Fail - Retry/Abort *)
IF _SubStep.isActive(_SUB_ADDRESS_RETRY_ABORT) THEN
	_retryAbort(
		numOfTargetRetries	:= _IparametersBase.numberOfRetries,
		retryAddress		:= _addressRestart, 
		abortAddress		:= _ADDRESS_FAIL);
END_IF
END_METHOD

METHOD PROTECTED _a2_X_KeyenceIVCameraTrigerDIO : BOOL 
VAR_INPUT
	camera					 : KOSTAL_AF2024_Drivers_Camera_I_Camera.I_CameraWithFeedback; 
	targetProgramNum		 : UINT;
	cameraName				 : STRING;
	
END_VAR
IF _step.toggle THEN 
	_stepDescription:= "TigerCameraKeyneceDIO";
END_IF

(* CheckCameraReady? *)
IF _SubStep.isActive(0) THEN 
	_addressRestart:= _SubStep.actual;
END_IF

(* Camera triger *)
IF _SubStep.isActive(1) THEN 
	IF NOT Camera.Ex_Trigger_ProgramNumber(ProgramNumber:= targetProgramNum) THEN 
		_updateHmiTextWithCameraBusy(name:= STRING_TO_WSTRING(cameraName));
	ELSIF NOT Camera.State.finish THEN 
		_updateHmiTextWithCameraBusy(name:= STRING_TO_WSTRING(cameraName));
	ELSIF NOT Camera.State.pass THEN 
		_getCameraErrorTexts(
			name		:= STRING_TO_WSTRING(cameraName),
			description	:= Camera.State.description);
		_a2_X_KeyenceIVCameraTrigerDIO:= FALSE;
	ELSE 
		_a2_X_KeyenceIVCameraTrigerDIO:= TRUE;
	END_IF
END_IF

//(* Pass *)
//IF _SubStep.isActive(_SUB_ADDRESS_PASS) THEN
//	_step.Condition:= TRUE;
//END_IF

//_step.Control();
END_METHOD

METHOD PROTECTED _a2_X_KeyenceIXCameraTriger : BOOL
VAR_INPUT
	Camera					 : TcNexa_Devices_Camera_TcCamera.I_Camera;
	IXtargerProgramNum	 	 : UINT;
	isIXcameraEnable		 : BOOL;
	IXcameraName			 : KOSTAL_AF2024_Core_Settings.T_MaxString_UTF8;
	
END_VAR
IF _step.toggle THEN 
	_stepDescription:= "IXCameraCheck";
END_IF

(*Chech parameters *)
IF _SubStep.isActive(0) THEN 
	IF NOT isIXcameraEnable THEN 
		_SubStep.set(request:= _SUB_ADDRESS_PASS);
	ELSE 
		_SubStep.INC();
	END_IF
END_IF
(* Set program number *)
IF _SubStep.isActive(0) THEN 
	Camera.setProgramNumber(
		programNumber:= IXtargerProgramNum,
		Response:= _InternalResponse);
	IF _InternalResponse.busy THEN 
		_updateHmiTextWithCameraBusy(name:= STRING_TO_WSTRING(IXcameraName));
	ELSE 
		_SubStep.INC(); 
	END_IF
END_IF 
(* Triger camera *)
IF _SubStep.isActive(2) THEN 
	Camera.inspect(Response:= _InternalResponse);
	IF _InternalResponse.busy THEN 
		_updateHmiTextWithCameraBusy(name:= STRING_TO_WSTRING( IXcameraName));
	ELSIF _InternalResponse.error THEN
//		_a2_X_KeyenceIXCameraTriger:= FALSE; 
		_getCameraErrorTexts(
			name:= STRING_TO_WSTRING(IXcameraName),
			description:= _Text.GetText(Number:= _E_TextCommon.camera_0_inError));
		_updateHmiText(
			userMessage:= STRING_TO_WSTRING( IXcameraName), 
			userAction:=  _Text.GetText(Number:= _E_TextCommon.camera_0_inError),
			isErrorMessage:= FALSE); 
	ELSE 
		_a2_X_KeyenceIXCameraTriger:= TRUE;
	END_IF
END_IF
(* Pass *)
IF _SubStep.isActive(_SUB_ADDRESS_PASS) THEN
	_step.Condition:= TRUE;
END_IF

_step.Control();
END_METHOD

METHOD PROTECTED _a2_X_KeyenceScanCode
VAR_INPUT
	Scanner				: KOSTAL_AF2024_Drivers_Scanner_IScanner.I_Scanner;
	isScannerEnable		: BOOL;
	ScannerName			: KOSTAL_AF2024_Core_Settings.T_MaxString;
END_VAR
VAR_OUTPUT
	SFC					: KOSTAL_AF2024_Core_Settings.T_MaxString_UTF8;
END_VAR
VAR 
	_tempInterger		: INT;
END_VAR
IF _step.toggle THEN 
	_stepDescription:= "ScanHousing";
	Scanner.ClearCodes();
END_IF

(* wait until scanner is ready *)
IF _SubStep.isActive(0) THEN 
	_addressRestart:= _SubStep.actual;
	IF NOT isScannerEnable THEN 
		_SubStep.set(request:= _SUB_ADDRESS_PASS);
		SFC:= '';
	ELSIF NOT Scanner.State.ready THEN 
		_Text.ClearVars();
		_Text.AddVar(Text:= ScannerName);
		_updateHmiText(
			userMessage		:= _Text.GetText(Number:= _E_TextCommon.scanner_0_failed),
			userAction		:= _Text.GetText(Number:= _E_TextCommon.scanner_0_notReady),
			isErrorMessage	:= FALSE);
	ELSE 
		_SubStep.INC();
	END_IF
END_IF
(* Execute *)
IF _SubStep.isActive(1) THEN 
	IF NOT Scanner.Ex_Scan() THEN 
		_Text.ClearVars();
		_Text.AddVar(Text:= ScannerName);
		_updateHmiText(
			userMessage		:= _Text.GetText(Number:= _E_TextCommon.scanner_0_busy),
			userAction		:= "",
			isErrorMessage	:= FALSE);	
	ELSIF NOT Scanner.State.finish THEN 
		_Text.ClearVars();
		_Text.AddVar(Text:= ScannerName);
		_updateHmiText(
			userMessage		:= _Text.GetText(Number:= _E_TextCommon.scanner_0_busy),
			userAction		:= "",
			isErrorMessage	:= FALSE);	
	ELSIF NOT Scanner.State.pass THEN 
		_Text.ClearVars();
		_Text.AddVar(Text:= ScannerName);
		_retryPartsInSeries:= _retryPartsInSeries+1 ;
		_subStepError:= _Text.GetText(Number:= _E_TextCommon.scanner_0_inError);
		_subStepMessage:= Scanner.State.description;
		_SubStep.set(request:= _SUB_ADDRESS_ABORT);
	ELSIF (Scanner.CodeGet(1) = '') OR (Scanner.CodeGet(1) = 'NONE') OR (Scanner.CodeGet(1) = 'Error') THEN 
		_Text.ClearVars();
		_Text.AddVar(Text:= ScannerName);
		_retryPartsInSeries:= _retryPartsInSeries+1 ;
			_subStepError:= _Text.GetText(Number:= _E_TextCommon.scanner_0_failed);
			_subStepMessage:= _Text.GetText(Number:= _E_TextCommon.barcodeNotfound);
			_SubStep.set(request:= _SUB_ADDRESS_RETRY_ABORT);
	ELSE 
		_SubStep.set(request:= _SUB_ADDRESS_PASS);
	END_IF
END_IF


(* Pass *)
IF _SubStep.isActive(_SUB_ADDRESS_PASS) THEN
	SFC:= Scanner.CodeGet(number:= 1);
	_step.Condition:= TRUE;
END_IF
(* Fail - Retry/Abort *)
IF _SubStep.isActive(_SUB_ADDRESS_RETRY_ABORT) THEN
	_retryAbort(
		numOfTargetRetries	:= _IparametersBase.numberOfRetries, 
		retryAddress		:= _addressRestart, 
		abortAddress		:= _ADDRESS_RUNOUT);
END_IF
(* Fail *)
IF _SubStep.isActive(_SUB_ADDRESS_ABORT) THEN
	_abort(abortAddress:= _ADDRESS_RUNOUT);
END_IF

_step.Control();
END_METHOD

METHOD PROTECTED _a2_X_LockPart
VAR_INPUT
	Cylinder		: KOSTAL_AF2024_Drivers_Actuation_Cylinder.I_Cylinder_Controlled;
END_VAR
IF _step.toggle THEN
	_stepDescription:= "LockHousing";
END_IF

(* Lock Housing *)
IF _SubStep.isActive(0) THEN
	IF Cylinder.moveTo_B() THEN
		_SubStep.set(request:= _SUB_ADDRESS_PASS);
	ELSIF Cylinder.Error.active THEN
		_subStepMessage:= Cylinder.Error.text;
		_SubStep.set(request:= _SUB_ADDRESS_RETRY_ABORT);
	ELSE
		_updateHmiTextWithCylinderTextMoveToWP(Cylinder:= Cylinder);
	END_IF
END_IF

(* Pass *)
IF _SubStep.isActive(_SUB_ADDRESS_PASS) THEN
	_step.Condition:= TRUE;
END_IF
(* Fail *)
IF _SubStep.isActive(_SUB_ADDRESS_RETRY_ABORT) THEN
	_retryAbort(
		numOfTargetRetries	:= _UNLIMITED_RETRY_NUMBER, 
		retryAddress		:= _addressRestart, 
		abortAddress		:= _ADDRESS_RUNOUT);
END_IF

_step.Control();
END_METHOD

METHOD PROTECTED _a2_X_PartNok
VAR_INPUT
END_VAR
IF _step.toggle THEN
	IF (_IresettableCounter <> 0) THEN _IresettableCounter.Fail.INC(); END_IF
	IF (_ItotalCounter <> 0) THEN _ItotalCounter.Fail.INC(); END_IF
	_partNok:= TRUE;
	_stepDescription:= "Part NOK";
	_subStepError:= "Part NOK";
	_subStepMessage:= "";
END_IF

_abort(abortAddress:= _ADDRESS_RUNOUT);
END_METHOD

METHOD PROTECTED _a2_X_PartOkWithCounter
VAR_INPUT
END_VAR
IF (_IresettableCounter <> 0) THEN _IresettableCounter.Pass.INC(); END_IF
IF (_ItotalCounter <> 0) THEN _ItotalCounter.Pass.INC(); END_IF
_partOk:= TRUE;
_step.set(request:= _ADDRESS_RUNOUT);
END_METHOD

METHOD PROTECTED _a2_X_PartOkWithoutCounter
VAR_INPUT
END_VAR
_partOk:= TRUE;
_step.set(request:= _ADDRESS_RUNOUT);
END_METHOD

METHOD PROTECTED _a2_X_RemovePart
VAR_INPUT
	partDetected		: BOOL;
END_VAR
IF _step.toggle THEN
	_stepDescription:= "RemovePart";
END_IF

IF _partOk THEN
	_updateHmiText(
		userMessage		:= _Text.GetText(Number:= _E_TextCommon.partOk),
		userAction		:= _Text.GetText(Number:= _E_TextCommon.removePart),
		isErrorMessage	:= FALSE);
ELSIF _partNok THEN
	_updateHmiText(
		userMessage		:= _Text.GetText(Number:= _E_TextCommon.partNok),
		userAction		:= _Text.GetText(Number:= _E_TextCommon.removePart),
		isErrorMessage	:= FALSE);
ELSE
	_updateHmiText(
		userMessage		:= _Text.GetText(Number:= _E_TextCommon.partUnknown),
		userAction		:= _Text.GetText(Number:= _E_TextCommon.removePart),
		isErrorMessage	:= FALSE);
END_IF

_step.Condition:= NOT partDetected;
_step.Control();
END_METHOD

METHOD PROTECTED _a2_X_TrigerCameraKeyenceTcpIp : BOOL
VAR_INPUT
	Camera					 : KOSTAL_AF2024_Drivers_Camera_Keyence_IV.I_Camera_TcpIp_IV;
	targerProgramNum		 : UINT;
	isCameraEnable			 : BOOL;
	cameraName				 : STRING;
	
END_VAR
IF _step.toggle THEN 
	_stepDescription:= "TigerCameraKeynece";
END_IF

(* CheckCameraReady? *)
IF _SubStep.isActive(0) THEN 
	_addressRestart:= _SubStep.actual;
	IF NOT isCameraEnable THEN 
//		_SubStep.set(request:= _SUB_ADDRESS_PASS);
		_a2_X_TrigerCameraKeyenceTcpIp:= TRUE;
	ELSIF NOT Camera.State.ready THEN 
		_updateHmiTextWithCameraNotReady(name:= STRING_TO_WSTRING (cameraName));
	ELSE 
		_SubStep.INC();
	END_IF
END_IF

(* Camera triger *)
IF _SubStep.isActive(1) THEN 
	IF NOT Camera.Ex_Trigger_ProgramNumber(ProgramNumber:= targerProgramNum) THEN 
		_updateHmiTextWithCameraBusy(name:= STRING_TO_WSTRING(cameraName));
	ELSIF NOT Camera.State.finish THEN 
		_updateHmiTextWithCameraBusy(name:= STRING_TO_WSTRING(cameraName));
	ELSIF NOT Camera.State.pass THEN 
		_a2_X_TrigerCameraKeyenceTcpIp:= FALSE;
		_getCameraErrorTexts(
			name		:= STRING_TO_WSTRING(cameraName),
			description	:= Camera.State.description);
		_SubStep.set(request:= _SUB_ADDRESS_RETRY_ABORT);
	ELSE 
//		_SubStep.set(request:= _SUB_ADDRESS_PASS);
		_a2_X_TrigerCameraKeyenceTcpIp:= TRUE;
	END_IF
END_IF

(* Pass *)
IF _SubStep.isActive(_SUB_ADDRESS_PASS) THEN
	_step.INC();
END_IF
(* Fail *)
IF _SubStep.isActive(_SUB_ADDRESS_RETRY_ABORT) THEN
	_retryAbort(
		numOfTargetRetries	:= _IparametersBase.numberOfRetries, 
		retryAddress		:= _addressRestart, 
		abortAddress		:= _ADDRESS_RUNOUT); //Check or address runout  ?
END_IF
END_METHOD

METHOD PROTECTED _a2_X_UnlockPart
VAR_INPUT
	Cylinder		: KOSTAL_AF2024_Drivers_Actuation_Cylinder.I_Cylinder_Controlled;
END_VAR
IF _step.toggle THEN
	_stepDescription:= "UnlockHousing";
END_IF

(* Unlock Housing *)
IF _SubStep.isActive(0) THEN
	IF Cylinder.moveTo_A() THEN
		_SubStep.set(request:= _SUB_ADDRESS_PASS);
	ELSIF Cylinder.Error.active THEN
		_addressRestart:= _SubStep.actual;
		_getCylinderErrorTexts(Cylinder:= Cylinder);
		_SubStep.set(request:= _SUB_ADDRESS_RETRY_ABORT);
	ELSE
		_updateHmiTextWithCylinderTextMoveToHP(Cylinder:= Cylinder);
	END_IF
END_IF
(* Pass *)
IF _SubStep.isActive(_SUB_ADDRESS_PASS) THEN
	_step.Condition:= TRUE;
END_IF
(* Fail *)
IF _SubStep.isActive(_SUB_ADDRESS_RETRY_ABORT) THEN
	_retryAbort(
		numOfTargetRetries	:= _UNLIMITED_RETRY_NUMBER, 
		retryAddress		:= _addressRestart, 
		abortAddress		:= _step.actual);
END_IF

_step.Control();
END_METHOD

METHOD PROTECTED _abort
VAR_INPUT
	abortAddress		: INT;
END_VAR
(* Abort button *)
_Hmi_station.Buttons_Custom.Button(7).Visible:= TRUE;
_Hmi_station.Buttons_Custom.Button(7).Text:= _Text.GetText(Number:= _E_TextCommon.abort);

_updateHmiText(
	userMessage		:= _subStepError, 
	userAction		:= _subStepMessage, 
	isErrorMessage	:= TRUE);

IF _Hmi_station.Buttons_Custom.Button(7).Pulse OR _IStation.pressedAbortButton  THEN //_onAbortButton.Q
	_condition.clear();
	_Hmi_station.Buttons_Custom.Button(7).Visible:= FALSE;
	_step.set(request:= abortAddress);
END_IF
END_METHOD

METHOD PROTECTED _checkCounterSPC
VAR_INPUT
END_VAR
IF _step.toggle THEN 
	_stepDescription:= "SpcCounterCheck";
END_IF

IF _SubStep.isActive(0) THEN 
	_counterForSCPmode:= _counterForSCPmode+1; 
	IF _counterForSCPmode > 5 THEN 
		_counterForSCPmode:= 0;
		_isSPCmodeActive:= FALSE;
		_step.set(request:= _ADDRESS_READY);
	ELSE 
		_isSPCmodeActive:= TRUE; 
		_SubStep.set(request:= _SUB_ADDRESS_PASS);
	END_IF
END_IF 

(* Pass *)
IF _SubStep.isActive(_SUB_ADDRESS_PASS) THEN
	_step.Condition:= TRUE;
END_IF

_step.Control();
END_METHOD

METHOD PROTECTED ABSTRACT _deviceDefine 
VAR_INPUT
END_VAR
END_METHOD

METHOD PROTECTED _getAxisErrorTexts
VAR_INPUT
	name 			: KOSTAL_AF2024_Core_Settings.T_MaxString;
	description		: KOSTAL_AF2024_Core_Settings.T_MaxString;
END_VAR
_Text.ClearVars();
_Text.AddVar(Text:= name);
_subStepError:= _Text.GetText(Number:= _E_TextCommon.axis_0_inError);
_subStepMessage:= description;
END_METHOD

METHOD PROTECTED _getCameraErrorTexts
VAR_INPUT
	name 			: KOSTAL_AF2024_Core_Settings.T_MaxString;
	description		: KOSTAL_AF2024_Core_Settings.T_MaxString;
END_VAR
_Text.ClearVars();
_Text.AddVar(Text:= name);
_subStepError:= _Text.GetText(Number:= _E_TextCommon.camera_0_failed);
_subStepMessage:= description;
END_METHOD

METHOD PROTECTED _getCameraIvToolResult : BOOL
VAR_INPUT
	Camera				: KOSTAL_AF2024_Drivers_Camera_Keyence_IV.I_Camera_TcpIp_IV;
	toolNum				: UDINT;
END_VAR
VAR
	_ICameraTool		: KOSTAL_AF2024_Drivers_Camera_Keyence_IV.I_T_Tool;
END_VAR
Camera.Result.Tools.Get_I(Number:= toolNum, rFound_I:= _ICameraTool, Response:= 0);
_getCameraIvToolResult:= _ICameraTool.Pass;
END_METHOD

METHOD PROTECTED _getCylinderErrorTexts
VAR_INPUT
	Cylinder			: KOSTAL_AF2024_Drivers_Actuation_Cylinder.I_Cylinder_Controlled;
END_VAR
_TextSplitter.Clear();
_TextSplitter.Split_Delimiter(
	Line		:= Cylinder.Name.device,
	Delimiter	:= "$L");
	
_Text.ClearVars();
_Text.AddVar(Text:= _TextSplitter.Results.line_GET(numberOfLine:= 1));
_subStepError:= _Text.GetText(Number:= _E_TextCommon.cylinder_0_inError);
_subStepMessage:= Cylinder.Error.text;
END_METHOD

METHOD PROTECTED _getLineControlErrorTexts
VAR_INPUT
	description		: KOSTAL_AF2024_Core_Settings.T_MaxString;
END_VAR
_Text.ClearVars();
_subStepError:= "Line Contorl failed";
_subStepMessage:= description;
END_METHOD

METHOD PROTECTED ABSTRACT _globalError
VAR_INPUT
END_VAR
END_METHOD

METHOD PROTECTED ABSTRACT _globalMessage
VAR_INPUT
END_VAR
END_METHOD

METHOD PROTECTED _handleCameraMaster
VAR_INPUT
	FirstShift 	: INT;
	SecondShift	: INT;
	ThirdShift	: INT;
END_VAR
VAR
	_tempTimeStruct		: Tc2_Utilities.TIMESTRUCT;
	_DT					: DATE_AND_TIME;
	_tempDint			: DINT;
	_isPreviousDay		: BOOL;
END_VAR
_onShiftChange(

	CLK:= 	(WORD_TO_INT(_IgetTime.TimeStruct.Hour) =   FirstShift)//6)

			OR ( WORD_TO_INT(_IgetTime.TimeStruct.Hour) =(SecondShift)) //14)

			OR ( WORD_TO_INT(_IgetTime.TimeStruct.Hour) = (ThirdShift)));//22));

IF _onShiftChange.Q OR NOT _cameraMasterOnStartupDone THEN 

	_IgetTime.TimeStruct.CopyTo(IN:= _tempTimeStruct); 

	_isPreviousDay := FALSE;

	IF (_tempTimeStruct.wHour >= INT_TO_WORD(FirstShift)) AND (_tempTimeStruct.wHour < INT_TO_WORD(SecondShift)) THEN 

		_tempTimeStruct.wHour:= INT_TO_WORD(FirstShift);

	ELSIF (_tempTimeStruct.wHour >= INT_TO_WORD(SecondShift)) AND (_tempTimeStruct.wHour < INT_TO_WORD(ThirdShift)) THEN 

		_tempTimeStruct.wHour:= INT_TO_WORD(SecondShift);

	ELSIF (_tempTimeStruct.wHour >= INT_TO_WORD(ThirdShift)) THEN

		_tempTimeStruct.wHour:= INT_TO_WORD(ThirdShift);

	ELSE 

		_tempTimeStruct.wHour:= INT_TO_WORD(ThirdShift);

		_isPreviousDay := TRUE;

	END_IF

	_tempTimeStruct.wMinute:= 0;

	_tempTimeStruct.wSecond:= 0;

	_tempTimeStruct.wMilliseconds:= 0;

	_DT:= Tc2_Utilities.SYSTEMTIME_TO_DT(TIMESTR:= _tempTimeStruct);

	_tempDint:= DT_TO_DINT(_DT);

	IF _isPreviousDay THEN

		_tempDint	:= _tempDint - 86400;

	END_IF

	IF (_tempDint > _lastCameraMasterTime) THEN 

		_isCameraMasterDone:= FALSE;
		_timeForMaster:= TRUE; 
		_lastCameraMasterTime:= _tempDint;

		_WritePersistentData(START:= TRUE);

	END_IF

	_cameraMasterOnStartupDone:= TRUE;

END_IF
 




//_onShiftChange(
//	CLK:= 	(WORD_TO_INT(_IgetTime.TimeStruct.Hour) =   FirstShift)//6)
//			OR ( WORD_TO_INT(_IgetTime.TimeStruct.Hour) =(SecondShift)) //14)
//			OR ( WORD_TO_INT(_IgetTime.TimeStruct.Hour) = (ThirdShift)));//22));
			
//IF _onShiftChange.Q OR NOT _cameraMasterOnStartupDone THEN 
//	_IgetTime.TimeStruct.CopyTo(IN:= _tempTimeStruct); 
//	IF (_tempTimeStruct.wHour >= INT_TO_WORD(FirstShift)) AND (_tempTimeStruct.wHour < INT_TO_WORD(SecondShift)) THEN 
//		_tempTimeStruct.wHour:= INT_TO_WORD(FirstShift);
//	ELSIF (_tempTimeStruct.wHour >= INT_TO_WORD(SecondShift)) AND (_tempTimeStruct.wHour < INT_TO_WORD(ThirdShift)) THEN 
//		_tempTimeStruct.wHour:= INT_TO_WORD(SecondShift);
//	ELSE 
//		_tempTimeStruct.wHour:= INT_TO_WORD(ThirdShift);
//	END_IF
//	_tempTimeStruct.wMinute:= 0;
//	_tempTimeStruct.wSecond:= 0;
//	_tempTimeStruct.wMilliseconds:= 0;
	
//	_DT:= Tc2_Utilities.SYSTEMTIME_TO_DT(TIMESTR:= _tempTimeStruct);
//	_tempDint:= DT_TO_DINT(_DT);
	
//	IF (_tempDint > _lastCameraMasterTime) THEN 
//		_isCameraMasterDone:= FALSE;
//		_lastCameraMasterTime:= _tempDint;
//		_WritePersistentData(START:= TRUE);
//	END_IF
	
//	_cameraMasterOnStartupDone:= TRUE;
//END_IF
END_METHOD

METHOD INTERNAL _handleCycleTime
VAR_INPUT
END_VAR
IF (_cycleTime <> _timerCycleTimer.ET) AND (_timerCycleTimer.ET <> T#0MS) THEN
	_cycleTime:= _timerCycleTimer.ET;
END_IF
END_METHOD

METHOD INTERNAL _handleManualModeStepDoneMessage
VAR_INPUT
END_VAR
IF _SubStep.isActive(stepNumber:= _SUB_ADDRESS_PASS) THEN
	_updateHmiText(
		userMessage		:= _Text.GetText(Number:= _E_TextCommon.stepDone),
		userAction		:= _Text.GetText(Number:= _E_TextCommon.stepContinue),
		isErrorMessage	:= FALSE);
END_IF
END_METHOD

METHOD _handlePersistentData
VAR_INPUT
END_VAR
_WritePersistentData(
	NETID	:= '',
	PORT	:= 851,
	START	:= FALSE,
	TMOUT	:= Tc2_System.DEFAULT_ADS_TIMEOUT);
END_METHOD

METHOD PROTECTED _handleProcessLight
VAR_INPUT
END_VAR
IF _mainControl.Mode.automatic THEN
	IF _partOk THEN
		DO_ProcessLightGreenLamp:= TRUE;
		DO_ProcessLightRedLamp:= FALSE;
		DO_ProcessLightYellowLamp:= FALSE;
		DO_ProcessLightBlueLamp:= FALSE;
	ELSIF _partNok THEN	
		DO_ProcessLightGreenLamp:= FALSE;
		DO_ProcessLightRedLamp:= TRUE;
		DO_ProcessLightYellowLamp:= FALSE;
		DO_ProcessLightBlueLamp:= FALSE;
	ELSIF _condition.isError() OR _condition.isMessage() THEN
		DO_ProcessLightGreenLamp:= FALSE;
		DO_ProcessLightRedLamp:= FALSE;
		DO_ProcessLightYellowLamp:= FALSE;
		DO_ProcessLightBlueLamp:= TRUE;	
	ELSE
		DO_ProcessLightGreenLamp:= FALSE;
		DO_ProcessLightRedLamp:= FALSE;
		DO_ProcessLightYellowLamp:= TRUE;
		DO_ProcessLightBlueLamp:= FALSE;	
	END_IF	
END_IF
END_METHOD

METHOD INTERNAL _hmiDefine
VAR
	_temp		: WSTRING;
END_VAR
_Hmi_station.FBmain();
(* Set station name *)
_temp:= TIME_TO_WSTRING(_cycleTime);
_temp:= Tc2_Standard.WRIGHT(
	STR:= _temp,
	SIZE:= Tc2_Standard.WLEN(_temp) - 2);
_Hmi_station.Name:= Tc2_Standard.WCONCAT(
	STR1:= _ID.name,
	STR2:= " [");
_Hmi_station.Name:= Tc2_Standard.WCONCAT(
	STR1:= _Hmi_station.Name,
	STR2:= _temp);
_Hmi_station.Name:= Tc2_Standard.WCONCAT(
	STR1:= _Hmi_station.Name,
	STR2:= "]");
_mainControl.ParticipantName:= _ID.name;
(* Set text lines on Hmi *)
_Hmi_station.Text.line_01:= _condition.Message.line_01;
_Hmi_station.Text.line_02:= _condition.Message.line_02;
_Hmi_station.Text.line_03:= _condition.Message.line_03;
_Hmi_station.Status.CopyFrom(IN:= _condition);
(* Reset button *)
_Hmi_station.Button_Escape.Visible:= _condition.isError() AND _mainControl.Mode.manual;
_Hmi_station.Button_Escape.Text:= _Text.GetText(Number:= _E_TextCommon.reset);
(* Plus button *)
_Hmi_station.Button_Plus.Visible:= _mainControl.Mode.manual AND (_step.actual > _ADDRESS_POWEROFF);
_Hmi_station.Button_Plus.Text:= _Text.GetText(Number:= _E_TextCommon.plus);
END_METHOD

METHOD INTERNAL _modeHandler
VAR_INPUT
END_VAR
_manualModeInterlock:= _mainControl.Mode.automatic OR NOT _state.Home;
_step.mode.automatic:= _mainControl.Mode.automatic AND NOT _condition.isError() AND NOT _cylinderInManualMode;
_step.mode.manual:= _mainControl.Mode.manual;
_step.StepNumberHome:= _ADDRESS_READY;
_step.LinkManual(
	Forward	:= _Hmi_station.Button_Plus.Pulse,
	Backward:= FALSE);
_step.ManualWithCondition:= TRUE;
END_METHOD

METHOD PROTECTED _moveCylinderToPossA : BOOL;
VAR_INPUT
	Cylinder			: I_Cylinder_Controlled;
END_VAR
IF Cylinder.moveTo_A() THEN 
	_moveCylinderToPossA:= TRUE;
ELSIF Cylinder.Error.active THEN 
	_moveCylinderToPossA:= FALSE;
	_updateHmiTextWithCylinderErrorSensorA(Cylinder:= Cylinder);
ELSE 
	_updateHmiTextWithCylinderTextMoveToHP(Cylinder:= Cylinder);
END_IF
END_METHOD

METHOD PROTECTED _moveCylinderToPossB : BOOL;
VAR_INPUT
	Cylinder			: I_Cylinder_Controlled;
END_VAR
IF Cylinder.moveTo_B() THEN 
	_moveCylinderToPossB:= TRUE;
ELSIF Cylinder.Error.active THEN 
	_moveCylinderToPossB:= FALSE;
	_updateHmiTextWithCylinderErrorSensorB(Cylinder:= Cylinder);
ELSE 
	_updateHmiTextWithCylinderTextMoveToWP(Cylinder:= Cylinder);
END_IF
END_METHOD

METHOD INTERNAL _resetCondition
VAR_INPUT
END_VAR
IF _condition.isError() THEN
	IF _Hmi_station.Button_Escape.Pulse THEN
		_condition.clear();
	END_IF
ELSE
	_condition.clear();	
END_IF
END_METHOD

METHOD INTERNAL _resetTcpIp
VAR_INPUT
END_VAR
_CloseAllSockets(bExecute:= NOT _isTcpIpInit);
_isTcpIpInit:= TRUE;
END_METHOD

METHOD PROTECTED _retryAbort
VAR_INPUT
	numOfTargetRetries	: INT;
	retryAddress		: INT;
	abortAddress		: INT;
END_VAR
(* Abort button *)
_Hmi_station.Buttons_Custom.Button(7).Visible:= TRUE;
_Hmi_station.Buttons_Custom.Button(7).Text:= _Text.GetText(Number:= _E_TextCommon.abort);
(* Retry button *)
IF (_retryPartsInSeries <= numOfTargetRetries) OR (numOfTargetRetries = _UNLIMITED_RETRY_NUMBER) THEN
	_Hmi_station.Buttons_Custom.Button(1).Visible:= TRUE;
	_Hmi_station.Buttons_Custom.Button(1).Text:= _Text.GetText(Number:= _E_TextCommon.retry);	
	_updateHmiText(
		userMessage		:= _subStepError, 
		userAction		:= _subStepMessage, 
		isErrorMessage	:= TRUE);
ELSE
	_Hmi_station.Buttons_Custom.Button(1).Visible:= FALSE;
	_updateHmiText(
		userMessage		:= _subStepError, 
		userAction		:= _subStepMessage,
		isErrorMessage	:= TRUE);
END_IF

IF (_Hmi_station.Buttons_Custom.Button(1).Pulse OR _onNagaraSwitch.Q) AND _Hmi_station.Buttons_Custom.Button(1).Visible THEN
	_condition.clear();
	_Hmi_station.Buttons_Custom.Button(1).Visible:= FALSE;
	_Hmi_station.Buttons_Custom.Button(7).Visible:= FALSE;
	_SubStep.set(request:= retryAddress);
ELSIF _Hmi_station.Buttons_Custom.Button(7).Pulse OR _IStation.pressedAbortButton THEN //_onAbortButton.Q 
	_condition.clear();
	_Hmi_station.Buttons_Custom.Button(1).Visible:= FALSE;
	_Hmi_station.Buttons_Custom.Button(7).Visible:= FALSE;
	_step.set(request:= abortAddress);
END_IF
END_METHOD

METHOD INTERNAL _stepHeader
VAR_INPUT
END_VAR
IF NOT _isStepInit THEN
	_step.init();
	_isStepInit:= TRUE;
ELSIF _mainControl.Demand.PowerOff AND (_step.actual <> _ADDRESS_POWEROFF) THEN
	_step.init();
END_IF

_step.Header();

(* Reset *)
IF _step.toggle THEN
	_stepDescription:= "";
	_Hmi_station.clear();
	_step.Condition:= FALSE;
	_step.JumpAddress:= 0;
	_SubStep.init();
	_retryPartsInSeries:= 0;
	_addressRestart:= 0;
END_IF
(* Sub step *)
IF (_lastSubStep <> _SubStep.actual) THEN
	_lastSubStep:= _SubStep.actual;
END_IF
END_METHOD

METHOD PROTECTED ABSTRACT _steps
VAR_INPUT
END_VAR
END_METHOD

METHOD PROTECTED _temepratureToleranceCheck  : BOOL
VAR_INPUT
	AnalogInput		: REAL;
	AnalogInputMin	: REAL;
	AnalogInputMax	: REAL;
END_VAR
IF AnalogInputMin < 0 THEN 
	IF AnalogInput < AnalogInputMin AND AnalogInput < AnalogInputMax THEN 
		_temepratureToleranceCheck:= TRUE;
	ELSE 
		_temepratureToleranceCheck:= FALSE;
	END_IF
ELSE 
	IF AnalogInput > AnalogInputMin AND AnalogInput < AnalogInputMax THEN 
		_temepratureToleranceCheck:= TRUE;
	ELSE 
		_temepratureToleranceCheck:= FALSE;
	END_IF
END_IF
END_METHOD

METHOD PROTECTED _TextReader : BOOL
VAR_INPUT
END_VAR
_Text.Path:= _TextPath;
_Text.FBmain();

IF _text.State.fail THEN
	_updateHmiText(
		userMessage		:= "TextHandler",
		userAction		:= _Text.State.description,
		isErrorMessage	:= TRUE);
ELSIF NOT _Text.Valid THEN
	_updateHmiText(
		userMessage		:= "TextHandler",
		userAction		:= _Text.State.description,
		isErrorMessage	:= FALSE);
END_IF

IF _text.LoadedLanguage <> '' THEN
	_textInitialized := TRUE;
END_IF
_TextReader := _textInitialized;
END_METHOD

METHOD PROTECTED _updateHmiText
VAR_INPUT
	userMessage		: KOSTAL_AF2024_Core_Settings.T_MaxString;
	userAction		: KOSTAL_AF2024_Core_Settings.T_MaxString;
	isErrorMessage	: BOOL;
END_VAR
_message.clear();

_Text.ClearVars();
_Text.AddVar(Text:= INT_TO_WSTRING(_step.actual));
_Text.AddVar(Text:= _stepDescription);
IF (_SubStep.actual = 32767) THEN
	_Text.AddVar(Text:= "0");	
ELSIF (_SubStep.actual <> _SUB_ADDRESS_ABORT) AND (_SubStep.actual <> _SUB_ADDRESS_RETRY_ABORT) THEN
	_Text.AddVar(Text:= INT_TO_WSTRING(_SubStep.actual));
ELSE
	_Text.AddVar(Text:= INT_TO_WSTRING(_lastSubStep));
END_IF
_message.line_01:= _Text.GetText(Number:= _E_TextCommon.step_0_actual_1);
_message.line_02:= userMessage;
_message.line_03:= userAction;
IF isErrorMessage AND NOT _condition.isError() THEN
	_log(Text:= _message.toString());
END_IF

IF isErrorMessage THEN
	_condition.setMessage(
		priority:= _condition.PriorityLevel_Error,
		message	:= _message);
ELSIF (userAction <> "") THEN
	_condition.setMessage(
		priority:= _condition.PriorityLevel_Message,
		message	:= _message);
ELSE
	_condition.setMessage(
		priority:= _condition.PriorityLevel_Text,
		message	:= _message);
END_IF
END_METHOD

METHOD PROTECTED _updateHmiTextWithAxisBusy
VAR_INPUT
	axisName			: KOSTAL_AF2024_Core_Settings.T_MaxString; 
END_VAR
_Text.ClearVars();
_Text.AddVar(Text:= axisName); 
_updateHmiText(
	userMessage		:=_Text.GetText(Number:= _E_TextCommon.axis_0_isBusy),
	userAction		:= "",
	isErrorMessage	:= FALSE);
END_METHOD

METHOD PROTECTED _updateHmiTextWithAxisNotReady
VAR_INPUT
END_VAR
_Text.ClearVars();
_updateHmiText(
	userMessage		:= _Text.GetText(Number:= _E_TextCommon.axis_0_notReady),
	userAction		:= "",
	isErrorMessage	:= FALSE);
END_METHOD

METHOD PROTECTED _updateHmiTextWithCameraBusy
VAR_INPUT
	name 			: KOSTAL_AF2024_Core_Settings.T_MaxString;
END_VAR
_Text.ClearVars();
_Text.AddVar(Text:= name);
_updateHmiText(
	userMessage		:= _Text.GetText(Number:= _E_TextCommon.camera_0_isBusy),
	userAction		:= "",
	isErrorMessage	:= FALSE);
END_METHOD

METHOD PROTECTED _updateHmiTextWithCameraNotReady
VAR_INPUT
	name		: KOSTAL_AF2024_Core_Settings.T_MaxString;
END_VAR
_Text.ClearVars();
_Text.AddVar(Text:= name);
_updateHmiText(
	userMessage		:= _Text.GetText(Number:= _E_TextCommon.camera_0_notReady),
	userAction		:= "",
	isErrorMessage	:= FALSE);
END_METHOD

METHOD PROTECTED _updateHmiTextWithCylinderError
VAR_INPUT
	Cylinder		: KOSTAL_AF2024_Drivers_Actuation_Cylinder.I_Cylinder_Controlled;
END_VAR
_TextSplitter.Clear();
_TextSplitter.Split_Delimiter(
	Line		:= Cylinder.Name.device,
	Delimiter	:=  "$L");

_Text.ClearVars();
_Text.AddVar(Text:= _TextSplitter.Results.line_GET(numberOfLine:= 1));
_updateHmiText(
	userMessage		:= _Text.GetText(Number:= _E_TextCommon.cylinder_0_inError),
	userAction		:= Cylinder.Error.text,
	isErrorMessage	:= TRUE);
_subStepError:= _Text.GetText(Number:= _E_TextCommon.cylinder_0_inError);
//_subStepMessage:= Cylinder.Error.text;

_TextSplitter.Split_Delimiter(
	Line		:= Cylinder.Name.sensor_A,
	Delimiter	:=  "$L");

_Text.AddVar(Text:= _TextSplitter.Results.line_GET(numberOfLine:= 2));
_subStepMessage:= _Text.GetText(Number:= _E_TextCommon.sensorFail);
END_METHOD

METHOD PROTECTED _updateHmiTextWithCylinderErrorSensorA
VAR_INPUT
	Cylinder		: KOSTAL_AF2024_Drivers_Actuation_Cylinder.I_Cylinder_Controlled;
END_VAR
_TextSplitter.Clear();
_TextSplitter.Split_Delimiter(
	Line		:= Cylinder.Name.device,
	Delimiter	:=  "$L");

_Text.ClearVars();
_Text.AddVar(Text:= _TextSplitter.Results.line_GET(numberOfLine:= 1));
_updateHmiText(
	userMessage		:= _Text.GetText(Number:= _E_TextCommon.cylinder_0_inError),
	userAction		:= Cylinder.Error.text,
	isErrorMessage	:= TRUE);
_subStepError:= _Text.GetText(Number:= _E_TextCommon.cylinder_0_inError);
//_subStepMessage:= Cylinder.Error.text;

_TextSplitter.Split_Delimiter(
	Line		:= Cylinder.Name.sensor_A,
	Delimiter	:=  "$L");

_Text.AddVar(Text:= _TextSplitter.Results.line_GET(numberOfLine:= 2));
_subStepMessage:= _Text.GetText(Number:= _E_TextCommon.sensorFail);
END_METHOD

METHOD PROTECTED _updateHmiTextWithCylinderErrorSensorB
VAR_INPUT
	Cylinder		: KOSTAL_AF2024_Drivers_Actuation_Cylinder.I_Cylinder_Controlled;
END_VAR
_TextSplitter.Clear();
_TextSplitter.Split_Delimiter(
	Line		:= Cylinder.Name.device,
	Delimiter	:=  "$L");

_Text.ClearVars();
_Text.AddVar(Text:= _TextSplitter.Results.line_GET(numberOfLine:= 1));
_updateHmiText(
	userMessage		:= _Text.GetText(Number:= _E_TextCommon.cylinder_0_inError),
	userAction		:= Cylinder.Error.text,
	isErrorMessage	:= TRUE);
_subStepError:= _Text.GetText(Number:= _E_TextCommon.cylinder_0_inError);
//_subStepMessage:= Cylinder.Error.text;

_TextSplitter.Split_Delimiter(
	Line		:= Cylinder.Name.sensor_B,
	Delimiter	:=  "$L");

_Text.AddVar(Text:= _TextSplitter.Results.line_GET(numberOfLine:= 2));
_subStepMessage:= _Text.GetText(Number:= _E_TextCommon.sensorFail);
END_METHOD

METHOD PROTECTED _updateHmiTextWithCylinderTextMoveToHP
VAR_INPUT
	Cylinder		: KOSTAL_AF2024_Drivers_Actuation_Cylinder.I_Cylinder_Controlled;
END_VAR
_TextSplitter.Clear();
_TextSplitter.Split_Delimiter(
	Line		:= Cylinder.Name.device,
	Delimiter	:=  "$L");

_Text.ClearVars();
_Text.AddVar(Text:= _TextSplitter.Results.line_GET(numberOfLine:= 1));
_updateHmiText(
	userMessage		:= _Text.GetText(Number:= _E_TextCommon.cylinder_0_moveToHPInProgress),
	userAction		:= "",
	isErrorMessage	:= FALSE);
_subStepError:= _Text.GetText(Number:= _E_TextCommon.cylinder_0_moveToHPInProgress);
_subStepMessage:= "";
END_METHOD

METHOD PROTECTED _updateHmiTextWithCylinderTextMoveToWP
VAR_INPUT
	Cylinder		: KOSTAL_AF2024_Drivers_Actuation_Cylinder.I_Cylinder_Controlled;
END_VAR
_TextSplitter.Clear();
_TextSplitter.Split_Delimiter(
	Line		:= Cylinder.Name.device,
	Delimiter	:=  "$L");

_Text.ClearVars();
_Text.AddVar(Text:= _TextSplitter.Results.line_GET(numberOfLine:= 1));
_updateHmiText(
	userMessage		:= _Text.GetText(Number:= _E_TextCommon.cylinder_0_moveToWPInProgress),
	userAction		:= "",
	isErrorMessage	:= FALSE);

_subStepError:= _Text.GetText(Number:= _E_TextCommon.cylinder_0_moveToWPInProgress);
_subStepMessage:= "";
END_METHOD

METHOD PROTECTED _updateHmiTextWithLineControlNotReady
VAR_INPUT
END_VAR
_Text.ClearVars();
_updateHmiText(
	userMessage:= "Line Contorl busy",
	userAction:= "",
	isErrorMessage:= FALSE);
END_METHOD

METHOD PROTECTED _updateHmiTextWithSensorFailText
VAR_INPUT
	sensorName		: KOSTAL_AF2024_Core_Settings.T_MaxString;
END_VAR
_Text.ClearVars();
_Text.AddVar(Text:= sensorName);
_updateHmiText(
	userMessage		:= _Text.GetText(Number:= _E_TextCommon.sensorFail),
	userAction		:= "",
	isErrorMessage	:= FALSE);
END_METHOD

METHOD FBmain
VAR_INPUT
END_VAR
IF NOT _parameterControl() THEN RETURN; END_IF

_onStateHome(CLK:= _state.Home);

_hmiDefine();
_resetTcpIp();
_deviceDefine();
_resetCondition();

IF NOT _TextReader() THEN RETURN; END_IF

_globalError();
_globalMessage();
_modeHandler();
_stepHeader();
_steps();
_handleProcessLight();
_handleCycleTime();
_handleManualModeStepDoneMessage();
//_handleCameraMaster(); //DA se definira lokalno ne vo baza
_handlePersistentData();
_onPowerOff(CLK:= _state.PowerOff);
_onNagaraSwitch(CLK:= DI_NagaraSwitch);
//_onAbortButton(CLK:= DI_AbortButton);
_onSubStepRetryAbort(CLK:= (_SubStep.actual = _SUB_ADDRESS_RETRY_ABORT));
IF _onSubStepRetryAbort.Q THEN
	_retryPartsInSeries:= _retryPartsInSeries + 1;
END_IF

_isDevicesInit:= TRUE;
END_METHOD

METHOD  linkCell
VAR_INPUT
	IN : I_CustomStationInterface; 
END_VAR
_IStation:= IN;
END_METHOD

END_FUNCTION_BLOCK

// ---- 03_FreeStations/03_TextMaster/DUTs/T_E_text_Common.TcPOU
FUNCTION_BLOCK T_E_text_Common EXTENDS KOSTAL_AF2024_Core_Text.T_E_Text
VAR
END_VAR

PROPERTY abort : KOSTAL_AF2024_Core_Text.ST_E_Text
GET
abort.Source:= KOSTAL_AF2024_Core_Text.E_Source.Common;
abort.Number:= 40;
END_GET
END_PROPERTY

PROPERTY axis_0_inError : KOSTAL_AF2024_Core_Text.ST_E_Text
GET
axis_0_inError.Source:= KOSTAL_AF2024_Core_Text.E_Source.Common;
axis_0_inError.Number:= 86;
END_GET
END_PROPERTY

PROPERTY axis_0_isBusy : KOSTAL_AF2024_Core_Text.ST_E_Text
GET
axis_0_isBusy.Source:= KOSTAL_AF2024_Core_Text.E_Source.Common;
axis_0_isBusy.Number:= 85;
END_GET
END_PROPERTY

PROPERTY axis_0_notReady : KOSTAL_AF2024_Core_Text.ST_E_Text
GET
axis_0_notReady.Source:= KOSTAL_AF2024_Core_Text.E_Source.Common;
axis_0_notReady.Number:= 87;
END_GET
END_PROPERTY

PROPERTY barcodeNotfound : KOSTAL_AF2024_Core_Text.ST_E_Text
GET
barcodeNotfound.Source:= KOSTAL_AF2024_Core_Text.E_Source.Common;
barcodeNotfound.Number:= 94;
END_GET
END_PROPERTY

PROPERTY camera_0_failed : KOSTAL_AF2024_Core_Text.ST_E_Text
GET
camera_0_failed.Source:= KOSTAL_AF2024_Core_Text.E_Source.Common;
camera_0_failed.Number:= 106;
END_GET
END_PROPERTY

PROPERTY camera_0_inError : KOSTAL_AF2024_Core_Text.ST_E_Text
GET
camera_0_inError.Source:= KOSTAL_AF2024_Core_Text.E_Source.Common;
camera_0_inError.Number:= 105;
END_GET
END_PROPERTY

PROPERTY camera_0_isBusy : KOSTAL_AF2024_Core_Text.ST_E_Text
GET
camera_0_isBusy.Source:= KOSTAL_AF2024_Core_Text.E_Source.Common;
camera_0_isBusy.Number:= 103;
END_GET
END_PROPERTY

PROPERTY camera_0_notReady : KOSTAL_AF2024_Core_Text.ST_E_Text
GET
camera_0_notReady.Source:= KOSTAL_AF2024_Core_Text.E_Source.Common;
camera_0_notReady.Number:= 104;
END_GET
END_PROPERTY

PROPERTY changeTool : KOSTAL_AF2024_Core_Text.ST_E_Text
GET
changeTool.Source:= KOSTAL_AF2024_Core_Text.E_Source.Common;
changeTool.Number:= 19;
END_GET
END_PROPERTY

PROPERTY clippingFailed : KOSTAL_AF2024_Core_Text.ST_E_Text
GET
clippingFailed.Source:= KOSTAL_AF2024_Core_Text.E_Source.Common;
clippingFailed.Number:= 20;
END_GET
END_PROPERTY

PROPERTY cylinder_0_inError : KOSTAL_AF2024_Core_Text.ST_E_Text
GET
cylinder_0_inError.Source:= KOSTAL_AF2024_Core_Text.E_Source.Common;
cylinder_0_inError.Number:= 82;
END_GET
END_PROPERTY

PROPERTY cylinder_0_moveToHPInProgress : KOSTAL_AF2024_Core_Text.ST_E_Text
GET
cylinder_0_moveToHPInProgress.Source:= KOSTAL_AF2024_Core_Text.E_Source.Common;
cylinder_0_moveToHPInProgress.Number:= 80;
END_GET
END_PROPERTY

PROPERTY cylinder_0_moveToWPInProgress : KOSTAL_AF2024_Core_Text.ST_E_Text
GET
cylinder_0_moveToWPInProgress.Source:= KOSTAL_AF2024_Core_Text.E_Source.Common;
cylinder_0_moveToWPInProgress.Number:= 81;
END_GET
END_PROPERTY

PROPERTY cylinderInManualMode : KOSTAL_AF2024_Core_Text.ST_E_Text
GET
cylinderInManualMode.Source:= KOSTAL_AF2024_Core_Text.E_Source.Common;
cylinderInManualMode.Number:= 52;
END_GET
END_PROPERTY

PROPERTY PUBLIC ExecutionNotAccepted : KOSTAL_AF2024_Core_Text.ST_E_Text
GET

ExecutionNotAccepted.Source:= Kostal_AF2024_Core_Text.E_Source.Common;
ExecutionNotAccepted.Number:= 117;
END_GET
END_PROPERTY

PROPERTY PUBLIC ExecutionNotFinished : KOSTAL_AF2024_Core_Text.ST_E_Text
GET

ExecutionNotFinished.Source:= Kostal_AF2024_Core_Text.E_Source.Common;
ExecutionNotFinished.Number:= 118;
END_GET
END_PROPERTY

PROPERTY firstCycle : KOSTAL_AF2024_Core_Text.ST_E_Text
GET
firstCycle.Source:= KOSTAL_AF2024_Core_Text.E_Source.Common;
firstCycle.Number:= 25;
END_GET
END_PROPERTY

PROPERTY insertMasterBadPart  : KOSTAL_AF2024_Core_Text.ST_E_Text
GET
insertMasterBadPart.Number:= 121;
END_GET
END_PROPERTY

PROPERTY insertMasterGoodPart  : KOSTAL_AF2024_Core_Text.ST_E_Text
GET
insertMasterGoodPart.Number:= 120;
END_GET
END_PROPERTY

PROPERTY insertPart : KOSTAL_AF2024_Core_Text.ST_E_Text
GET
insertPart.Source:= KOSTAL_AF2024_Core_Text.E_Source.Common;
insertPart.Number:= 61;
END_GET
END_PROPERTY

PROPERTY lastCycle : KOSTAL_AF2024_Core_Text.ST_E_Text
GET
lastCycle.Source:= KOSTAL_AF2024_Core_Text.E_Source.Common;
lastCycle.Number:= 27;
END_GET
END_PROPERTY

PROPERTY mainControlIsIn_0_state : KOSTAL_AF2024_Core_Text.ST_E_Text
GET
mainControlIsIn_0_state.Source:= KOSTAL_AF2024_Core_Text.E_Source.Common;
mainControlIsIn_0_state.Number:= 10;
END_GET
END_PROPERTY

PROPERTY noArticleSelected : KOSTAL_AF2024_Core_Text.ST_E_Text
GET
noArticleSelected.Source:= KOSTAL_AF2024_Core_Text.E_Source.Common;
noArticleSelected.Number:= 17;
END_GET
END_PROPERTY

PROPERTY normalCycle : KOSTAL_AF2024_Core_Text.ST_E_Text
GET
normalCycle.Source:= KOSTAL_AF2024_Core_Text.E_Source.Common;
normalCycle.Number:= 26;
END_GET
END_PROPERTY

PROPERTY off : KOSTAL_AF2024_Core_Text.ST_E_Text
GET
off.Source:= KOSTAL_AF2024_Core_Text.E_Source.Common;
off.Number:= 2;
END_GET
END_PROPERTY

PROPERTY on : KOSTAL_AF2024_Core_Text.ST_E_Text
GET
on.Source:= KOSTAL_AF2024_Core_Text.E_Source.Common;
on.Number:= 3;
END_GET
END_PROPERTY

PROPERTY partNok : KOSTAL_AF2024_Core_Text.ST_E_Text
GET
partNok.Source:= KOSTAL_AF2024_Core_Text.E_Source.Common;
partNok.Number:= 55;
END_GET
END_PROPERTY

PROPERTY partOk : KOSTAL_AF2024_Core_Text.ST_E_Text
GET
partOk.Source:= KOSTAL_AF2024_Core_Text.E_Source.Common;
partOk.Number:= 54;
END_GET
END_PROPERTY

PROPERTY partUnknown : KOSTAL_AF2024_Core_Text.ST_E_Text
GET
partUnknown.Source:= KOSTAL_AF2024_Core_Text.E_Source.Common;
partUnknown.Number:= 56;
END_GET
END_PROPERTY

PROPERTY plus : KOSTAL_AF2024_Core_Text.ST_E_Text
GET
plus.Source:= Kostal_AF2024_Core_Text.E_Source.Common;
plus.Number:= 6;
END_GET
END_PROPERTY

PROPERTY pressNagara : KOSTAL_AF2024_Core_Text.ST_E_Text
GET
pressNagara.Source:= KOSTAL_AF2024_Core_Text.E_Source.Common;
pressNagara.Number:= 60;
END_GET
END_PROPERTY

PROPERTY printer_0_inError : KOSTAL_AF2024_Core_Text.ST_E_Text
GET
printer_0_inError.Number:= 110;
END_GET
END_PROPERTY

PROPERTY printer_0_isBusy  : KOSTAL_AF2024_Core_Text.ST_E_Text
GET
printer_0_isBusy.Number:= 108;
END_GET
END_PROPERTY

PROPERTY printer_0_notReady  : KOSTAL_AF2024_Core_Text.ST_E_Text
GET
printer_0_notReady.Number:= 109;
END_GET
END_PROPERTY

PROPERTY removePart : KOSTAL_AF2024_Core_Text.ST_E_Text
GET
removePart.Source:= KOSTAL_AF2024_Core_Text.E_Source.Common;
removePart.Number:= 57;
END_GET
END_PROPERTY

PROPERTY reset : KOSTAL_AF2024_Core_Text.ST_E_Text
GET
reset.Source:= Kostal_AF2024_Core_Text.E_Source.Common;
reset.Number:= 7;
END_GET
END_PROPERTY

PROPERTY retry : KOSTAL_AF2024_Core_Text.ST_E_Text
GET
retry.Source:= KOSTAL_AF2024_Core_Text.E_Source.Common;
retry.Number:= 41;
END_GET
END_PROPERTY

PROPERTY scanner_0_busy : KOSTAL_AF2024_Core_Text.ST_E_Text
GET
scanner_0_busy.Source:= KOSTAL_AF2024_Core_Text.E_Source.Common;
scanner_0_busy.Number:= 90;
END_GET
END_PROPERTY

PROPERTY scanner_0_failed : KOSTAL_AF2024_Core_Text.ST_E_Text
GET
scanner_0_failed.Source:= KOSTAL_AF2024_Core_Text.E_Source.Common;
scanner_0_failed.Number:= 93;
END_GET
END_PROPERTY

PROPERTY scanner_0_inError : KOSTAL_AF2024_Core_Text.ST_E_Text
GET
scanner_0_inError.Source:= KOSTAL_AF2024_Core_Text.E_Source.Common;
scanner_0_inError.Number:= 92;
END_GET
END_PROPERTY

PROPERTY scanner_0_noCode : KOSTAL_AF2024_Core_Text.ST_E_Text
GET
scanner_0_noCode.Source:= KOSTAL_AF2024_Core_Text.E_Source.Common;
scanner_0_noCode.Number:= 94;
END_GET
END_PROPERTY

PROPERTY scanner_0_notReady : KOSTAL_AF2024_Core_Text.ST_E_Text
GET
scanner_0_notReady.Source:= KOSTAL_AF2024_Core_Text.E_Source.Common;
scanner_0_notReady.Number:= 91;
END_GET
END_PROPERTY

PROPERTY selectArticle : KOSTAL_AF2024_Core_Text.ST_E_Text
GET
selectArticle.Source:= KOSTAL_AF2024_Core_Text.E_Source.Common;
selectArticle.Number:= 18;
END_GET
END_PROPERTY

PROPERTY sensorFail : KOSTAL_AF2024_Core_Text.ST_E_Text
GET
sensorFail.Source:= Kostal_AF2024_Core_Text.E_Source.Common;
sensorFail.Number:= 70;
END_GET
END_PROPERTY

PROPERTY sensorOverlap : KOSTAL_AF2024_Core_Text.ST_E_Text
GET
sensorOverlap.Source:= Kostal_AF2024_Core_Text.E_Source.Common;
sensorOverlap.Number:= 71;
END_GET
END_PROPERTY

PROPERTY sliderPullOut : KOSTAL_AF2024_Core_Text.ST_E_Text
GET
sliderPullOut.Source:= KOSTAL_AF2024_Core_Text.E_Source.Common;
sliderPullOut.Number:= 67;
END_GET
END_PROPERTY

PROPERTY sliderPushIn : KOSTAL_AF2024_Core_Text.ST_E_Text
GET
sliderPushIn.Source:= KOSTAL_AF2024_Core_Text.E_Source.Common;
sliderPushIn.Number:= 68;
END_GET
END_PROPERTY

PROPERTY start : KOSTAL_AF2024_Core_Text.ST_E_Text
GET
start.Source:= KOSTAL_AF2024_Core_Text.E_Source.Common;
start.Number:= 5;
END_GET
END_PROPERTY

PROPERTY stationInManualMode : KOSTAL_AF2024_Core_Text.ST_E_Text
GET
stationInManualMode.Source:= KOSTAL_AF2024_Core_Text.E_Source.Common;
stationInManualMode.Number:= 51;
END_GET
END_PROPERTY

PROPERTY stationReady : KOSTAL_AF2024_Core_Text.ST_E_Text
GET
stationReady.Source:= KOSTAL_AF2024_Core_Text.E_Source.Common;
stationReady.Number:= 50;
END_GET
END_PROPERTY

PROPERTY step_0_actual_1 : KOSTAL_AF2024_Core_Text.ST_E_Text
GET
step_0_actual_1.Source:= KOSTAL_AF2024_Core_Text.E_Source.Common;
step_0_actual_1.Number:= 11;
END_GET
END_PROPERTY

PROPERTY step_0_doesNotExist : KOSTAL_AF2024_Core_Text.ST_E_Text
GET
step_0_doesNotExist.Source:= KOSTAL_AF2024_Core_Text.E_Source.Common;
step_0_doesNotExist.Number:= 12;
END_GET
END_PROPERTY

PROPERTY stepContinue : KOSTAL_AF2024_Core_Text.ST_E_Text
GET
stepContinue.Source:= KOSTAL_AF2024_Core_Text.E_Source.Common;
stepContinue.Number:= 14;
END_GET
END_PROPERTY

PROPERTY stepDone : KOSTAL_AF2024_Core_Text.ST_E_Text
GET
stepDone.Source:= KOSTAL_AF2024_Core_Text.E_Source.Common;
stepDone.Number:= 13;
END_GET
END_PROPERTY

PROPERTY stop : KOSTAL_AF2024_Core_Text.ST_E_Text
GET
stop.Source:= KOSTAL_AF2024_Core_Text.E_Source.Common;
stop.Number:= 4;
END_GET
END_PROPERTY

PROPERTY unknownProductType : KOSTAL_AF2024_Core_Text.ST_E_Text
GET
unknownProductType.Source:= KOSTAL_AF2024_Core_Text.E_Source.Common;
unknownProductType.Number:= 115;
END_GET
END_PROPERTY

PROPERTY valveNotOn : KOSTAL_AF2024_Core_Text.ST_E_Text
GET
valveNotOn.Number:= 73;
END_GET
END_PROPERTY

PROPERTY waitForSensor_0 : KOSTAL_AF2024_Core_Text.ST_E_Text
GET
waitForSensor_0.Source:= KOSTAL_AF2024_Core_Text.E_Source.Common;
waitForSensor_0.Number:= 72;
END_GET
END_PROPERTY

PROPERTY waitSliderInBackPosition : KOSTAL_AF2024_Core_Text.ST_E_Text
GET
waitSliderInBackPosition.Source:= KOSTAL_AF2024_Core_Text.E_Source.Common;
waitSliderInBackPosition.Number:= 66;
END_GET
END_PROPERTY

PROPERTY waitSliderInFrontPosition : KOSTAL_AF2024_Core_Text.ST_E_Text
GET
waitSliderInFrontPosition.Source:= KOSTAL_AF2024_Core_Text.E_Source.Common;
waitSliderInFrontPosition.Number:= 65;
END_GET
END_PROPERTY

PROPERTY wrongLowerTool : KOSTAL_AF2024_Core_Text.ST_E_Text
GET
wrongLowerTool.Source:= KOSTAL_AF2024_Core_Text.E_Source.Common;
wrongLowerTool.Number:= 15;
END_GET
END_PROPERTY

PROPERTY wrongUpperTool : KOSTAL_AF2024_Core_Text.ST_E_Text
GET
wrongUpperTool.Source:= KOSTAL_AF2024_Core_Text.E_Source.Common;
wrongUpperTool.Number:= 16;
END_GET
END_PROPERTY

END_FUNCTION_BLOCK

// ---- 02_ControlledStations/FB_StationBaseWithAutomaticSlider.TcPOU
FUNCTION_BLOCK ABSTRACT FB_StationBaseWithAutomaticSlider EXTENDS FB_StationBase
VAR
	(* Slider Automatic Cylinder *)
	_SliderAutomaticCylinder 				   : KOSTAL_AF2024_Drivers_Actuation_Cylinder.FB_Cylinder_Controlled;
	DI_SliderAutomaticCylinderHP		AT %I* : BOOL;
	DI_SliderAutomaticCylinderWP		AT %I* : BOOL;
	DO_SliderAutomaticCylinderWP		AT %Q* : BOOL;
	DO_SliderAutomaticCylinderHP		AT %Q* : BOOL;
	
	(* Slider Locking Cylinder Front Position *)
	_SliderLockingCylinderFrontPosition		: KOSTAL_AF2024_Drivers_Actuation_Cylinder.FB_Cylinder_Controlled;
	DO_SliderLockCylinderFrontPosHP		AT %Q* : BOOL; // Treba da se vidi koi sensori bi se koristele ovde 
	DO_SliderLockCylinderFrontPosWP		AT %Q* : BOOL;
	DI_SliderLockCylinderFrontPosWP		AT %I* : BOOL;
	DI_SliderLockCylinderFrontPosHP		AT %I* : BOOL;
	DI_SliderInFrontPos					AT %I* : BOOL;
	DI_SliderInBackPos					AT %I* : BOOL;
	
	(* Process *)
	_timerSliderInBackPos						: Tc2_Standard.TON;
	_timerSliderInFrontPos						: Tc2_Standard.TON;
	
	(* Names *)
	_automaticSliderInFrontPositionName 	: KOSTAL_AF2024_Core_Settings.T_MaxString;
	_automaticSliderInBackPositionName 	: KOSTAL_AF2024_Core_Settings.T_MaxString;
	_isHomeDone					: BOOL;
END_VAR

METHOD PROTECTED _a2_X_CloseAutomaticSlider
VAR_INPUT
END_VAR
IF _step.toggle THEN
	_timerSliderInFrontPos(IN:= FALSE);
	_stepDescription:= "SliderUnlockFrontPosition"; 
END_IF

(* If slider in front position skip this step *)
IF _SubStep.isActive(0) THEN 
	IF DI_SliderAutomaticCylinderWP THEN 
		_SubStep.set(request:= 4);
	ELSE 
		_SubStep.INC();
	END_IF
END_IF 
(* Unlock *)
IF _SubStep.isActive(1) THEN 
	IF _SliderLockingCylinderFrontPosition.moveTo_A() THEN 
		_SubStep.INC();
	ELSIF  _SliderLockingCylinderFrontPosition.Error.active THEN 	
		_updateHmiTextWithCylinderError(Cylinder:= _SliderLockingCylinderFrontPosition);
		_SubStep.set(request:= _SUB_ADDRESS_RETRY_ABORT);
	ELSE 
		_updateHmiTextWithCylinderTextMoveToHP(Cylinder:= _SliderLockingCylinderFrontPosition);
	END_IF
END_IF
(* Move Automatic Slider Cylinder in front position*)
IF _SubStep.isActive(2) THEN 
	IF _SliderAutomaticCylinder.moveTo_B() THEN 
		_SubStep.INC();
	ELSIF _SliderAutomaticCylinder.Error.active THEN 
		_updateHmiTextWithCylinderError(Cylinder:= _SliderAutomaticCylinder);
	ELSE 
		_updateHmiTextWithCylinderTextMoveToWP(Cylinder:= _SliderAutomaticCylinder);
	END_IF
END_IF
(* Wait slider in back position *)
IF _SubStep.isActive(3) THEN 
	_timerSliderInFrontPos(
		IN	:= DI_SliderAutomaticCylinderWP,
		PT	:= T#500MS); //T#500MS
	IF NOT _timerSliderInFrontPos.Q THEN  
		_Text.ClearVars();
		_Text.AddVar(Text:= _automaticSliderInFrontPositionName);
		_updateHmiText(
			userMessage		:= _Text.GetText(Number:= _E_TextCommon.waitSliderInFrontPosition),
			userAction		:= _Text.GetText(Number:= _E_TextCommon.waitForSensor_0),
			isErrorMessage	:= FALSE);	
	ELSIF  DI_SliderAutomaticCylinderWP  THEN 
		_SubStep.INC();
	END_IF	
END_IF
(* Lock *)
IF _SubStep.isActive(4) THEN
	IF _SliderLockingCylinderFrontPosition.moveTo_B() THEN
		_SliderAutomaticCylinder.Pressureless();
		_SubStep.set(request:= _SUB_ADDRESS_PASS);
	ELSIF _SliderLockingCylinderFrontPosition.Error.active THEN
		_addressRestart:= _SubStep.actual;
		_getCylinderErrorTexts(Cylinder:= _SliderLockingCylinderFrontPosition);
		_SubStep.set(request:= _SUB_ADDRESS_RETRY_ABORT);
	ELSE
		_updateHmiTextWithCylinderTextMoveToWP(Cylinder:= _SliderLockingCylinderFrontPosition);
	END_IF
END_IF
(* Pass *)
IF _SubStep.isActive(_SUB_ADDRESS_PASS) THEN
	_step.Condition:= TRUE;
END_IF
(* Fail *)
IF _SubStep.isActive(_SUB_ADDRESS_RETRY_ABORT) THEN
	_retryAbort(
		numOfTargetRetries	:= _UNLIMITED_RETRY_NUMBER,
		retryAddress		:= _addressRestart,
		abortAddress		:= _ADDRESS_RUNOUT);
END_IF

_step.Control();
END_METHOD

METHOD PROTECTED _a2_X_OpenAutomaticSlider
VAR_INPUT
END_VAR
IF _step.toggle THEN 
	_timerSliderInBackPos(IN:= FALSE);
	_stepDescription:= "CloseAutomaticSlider";
END_IF
(* If slider in back position skip this step *)
IF _SubStep.isActive(0) THEN 
	IF DI_SliderAutomaticCylinderHP THEN 
		_SubStep.set(request:=3);
	ELSE 
		_SubStep.INC();
	END_IF
END_IF 
(* Unlock *)
IF _SubStep.isActive(1) THEN 
	IF _SliderLockingCylinderFrontPosition.moveTo_A() THEN 
		_SubStep.INC();
	ELSIF  _SliderLockingCylinderFrontPosition.Error.active THEN 
		_updateHmiTextWithCylinderError(Cylinder:= _SliderLockingCylinderFrontPosition);
		_SubStep.set(request:= _SUB_ADDRESS_RETRY_ABORT);
	ELSE 
		_updateHmiTextWithCylinderTextMoveToHP(Cylinder:= _SliderLockingCylinderFrontPosition);
	END_IF
END_IF
(* Move Automatic Slider Cylinder in back position*)
IF _SubStep.isActive(2) THEN 
	IF _SliderAutomaticCylinder.moveTo_A() THEN 
		_SubStep.INC();
	ELSIF _SliderAutomaticCylinder.Error.active THEN 
		_updateHmiTextWithCylinderError(Cylinder:= _SliderAutomaticCylinder);
	ELSE 
		_updateHmiTextWithCylinderTextMoveToWP(Cylinder:= _SliderAutomaticCylinder);
	END_IF
END_IF
(* Wait slider in back position *)
IF _SubStep.isActive(3) THEN 
	_timerSliderInBackPos(
		IN:=   DI_SliderAutomaticCylinderHP,
		PT:=   T#500MS 	);//500ms da se doddade
	IF NOT DI_SliderAutomaticCylinderHP THEN 
		_Text.ClearVars();
		_Text.AddVar(Text:= _automaticSliderInBackPositionName);
		_updateHmiText(
			userMessage		:= _Text.GetText(Number:= _E_TextCommon.waitSliderInBackPosition),
			userAction		:= _Text.GetText(Number:= _E_TextCommon.waitForSensor_0),
			isErrorMessage	:= FALSE);
	ELSIF NOT _timerSliderInBackPos.Q THEN 
		_Text.ClearVars();
		_Text.AddVar(Text:= _automaticSliderInBackPositionName);
		_updateHmiText(
			userMessage		:= _Text.GetText(Number:= _E_TextCommon.waitSliderInBackPosition),
			userAction		:= _Text.GetText(Number:= _E_TextCommon.waitForSensor_0),
			isErrorMessage	:= FALSE);	
	ELSE 
		_SubStep.set(request:= _SUB_ADDRESS_PASS);
	END_IF	
END_IF
//(* Lock *)
//IF _SubStep.isActive(4) THEN
//	IF _SliderLockingCylinderFrontPosition.moveTo_B() THEN
//		_SubStep.set(request:= _SUB_ADDRESS_PASS);
//	ELSIF _SliderLockingCylinderFrontPosition.Error.active THEN
//		_addressRestart:= _SubStep.actual;
//		_getCylinderErrorTexts(Cylinder:= _SliderLockingCylinderFrontPosition);
//		_SubStep.set(request:= _SUB_ADDRESS_RETRY_ABORT);
//	ELSE
//		_updateHmiTextWithCylinderTextMoveToWP(Cylinder:= _SliderLockingCylinderFrontPosition);
//	END_IF
//END_IF
(* Pass *)
IF _SubStep.isActive(_SUB_ADDRESS_PASS) THEN
	_step.Condition:= TRUE;
END_IF
(* Fail *)
IF _SubStep.isActive(_SUB_ADDRESS_RETRY_ABORT) THEN
	_retryAbort(
		numOfTargetRetries	:= _UNLIMITED_RETRY_NUMBER,
		retryAddress		:= _addressRestart,
		abortAddress		:= _ADDRESS_RUNOUT);
END_IF

_step.Control();
END_METHOD

PROPERTY sliderInBackPositionName : KOSTAL_AF2024_Core_Settings.T_MaxString
GET
sliderInBackPositionName:= _automaticSliderInBackPositionName;
END_GET
SET
_automaticSliderInBackPositionName:= sliderInBackPositionName;
END_SET
END_PROPERTY

PROPERTY sliderInFrontPositionName : KOSTAL_AF2024_Core_Settings.T_MaxString
GET
sliderInFrontPositionName:= _automaticSliderInFrontPositionName;
END_GET
SET
_automaticSliderInFrontPositionName:= sliderInFrontPositionName;
END_SET
END_PROPERTY

END_FUNCTION_BLOCK

// ---- 02_ControlledStations/FB_StationBaseWithSlider.TcPOU
FUNCTION_BLOCK ABSTRACT FB_StationBaseWithSlider EXTENDS FB_StationBase
VAR
	(* General *)
	_IparametersCommon						: I_Parameters_MainControl;
	(* Slider Lock Cylinder *)    	
	_SliderLockCylinderInFrontPosition		: KOSTAL_AF2024_Drivers_Actuation_Cylinder.FB_Cylinder_Controlled;	

	DI_SliderInFrontPos						AT %I* : BOOL;
	DI_SliderInBackPos						AT %I* : BOOL;
	DI_SliderLockCylInFrontPosWP			AT %I* : BOOL;
	DI_SliderLockCylInFrontPosHP			AT %I* : BOOL;
	DO_SliderLockCylInFrontPosHP			AT %Q* : BOOL;
	DO_SliderLockCylInFrontPosWP			AT %Q* : BOOL;	  
	
	(* Sensors *)
	_sliderInFrontPositionName 	: KOSTAL_AF2024_Core_Settings.T_MaxString;
	_sliderInBackPositionName 	: KOSTAL_AF2024_Core_Settings.T_MaxString;
	(* Process *)
	_timerSliderInFrontPos		: Tc2_Standard.TON;
	_timerSliderInBackPos		: Tc2_Standard.TON;
	
	(* Axis *)
//	_Axis						: KOSTAL_TC3_Device_Axis_FESTO_CMMT_AS_ETC.FB_FESTO_CMMT_AS;
	_isHomeDone					: BOOL;
//	_AxisName					: KOSTAL_AF2024_Core_Settings.T_MaxString;
	
END_VAR

METHOD _a2_X_CloseSlider
VAR_INPUT
END_VAR
IF _step.toggle THEN 
	_timerSliderInBackPos(IN:= FALSE);
	_stepDescription:= "CloseSlider";
END_IF

(* If slider in back position skip this step *)
IF _SubStep.isActive(0) THEN 
	_timerSliderInBackPos(IN:= FALSE);
	_addressRestart:= _SubStep.actual;
	IF DI_SliderInBackPos THEN 
		_SubStep.set(request:= 3);
	ELSE 
		_SubStep.INC();
	END_IF
END_IF 

(* Unlock *)
IF _SubStep.isActive(1) THEN 
	IF _SliderLockCylinderInFrontPosition.moveTo_B() THEN 
		_SubStep.INC();
	ELSIF _SliderLockCylinderInFrontPosition.Error.active THEN 
		_addressRestart:= _SubStep.actual;
		_getCylinderErrorTexts(Cylinder:= _SliderLockCylinderInFrontPosition);
		_SubStep.set(request:= _SUB_ADDRESS_RETRY_ABORT);
	ELSE 
		_updateHmiTextWithCylinderTextMoveToHP(Cylinder:= _SliderLockCylinderInFrontPosition);
	END_IF
END_IF

(* Wait sluder in back position *)
IF _SubStep.isActive(2) THEN 
	_timerSliderInBackPos(
		IN 	:= DI_SliderInBackPos,
		PT	:= T#150MS);
	IF NOT DI_SliderInBackPos THEN 
		_Text.ClearVars();
		_Text.AddVar(Text:= _sliderInBackPositionName);
		_updateHmiText(
			userMessage		:= _Text.GetText(Number:= _E_TextCommon.waitSliderInBackPosition),
			userAction		:= _Text.GetText(Number:= _E_TextCommon.waitForSensor_0),
			isErrorMessage	:= FALSE);
	ELSIF _timerSliderInBackPos.Q THEN 
		_SubStep.INC();
	END_IF
END_IF 

(* Lock slider in back position *)
IF _SubStep.isActive(3) THEN
	DO_SliderLockCylInFrontPosWP:= FALSE; 
	IF  _SliderLockCylinderInFrontPosition.moveTo_A()   THEN
		_SubStep.set(request:= _SUB_ADDRESS_PASS);
	ELSIF _SliderLockCylinderInFrontPosition.Error.active THEN
		_getCylinderErrorTexts(Cylinder:= _SliderLockCylinderInFrontPosition);
		_SubStep.set(request:= _SUB_ADDRESS_RETRY_ABORT);
	ELSE
		_updateHmiTextWithCylinderTextMoveToWP(Cylinder:= _SliderLockCylinderInFrontPosition);
	END_IF
END_IF
(* Pass *)
IF _SubStep.isActive(_SUB_ADDRESS_PASS) THEN
	_step.Condition:= TRUE;
END_IF
(* Fail *)
IF _SubStep.isActive(_SUB_ADDRESS_RETRY_ABORT) THEN
	_retryAbort(
		numOfTargetRetries	:= _UNLIMITED_RETRY_NUMBER,
		retryAddress		:= _addressRestart,
		abortAddress		:= _ADDRESS_RUNOUT); //?
END_IF

_step.Control();
END_METHOD

METHOD PROTECTED _a2_X_HomeAxes
VAR_INPUT
	axis1			: REFERENCE TO  KOSTAL_AF2024_Drivers_Actuation_Axis_Festo_CMMT_AS.FB_FESTO_CMMT_AS;
	axisName1		: KOSTAL_AF2024_Core_Settings.T_MaxString;
	axis2			: REFERENCE TO  KOSTAL_AF2024_Drivers_Actuation_Axis_Festo_CMMT_AS.FB_FESTO_CMMT_AS;
	axisName2		: KOSTAL_AF2024_Core_Settings.T_MaxString;
END_VAR
 IF _step.toggle THEN 
	_stepDescription:= "HomeAxis";
END_IF

(* Home axis Left*)
IF _SubStep.isActive(0) THEN 
	 IF NOT axis1.Ex_Homing() THEN
		 _updateHmiTextWithAxisBusy(axisName:= axisName1);		 
	ELSIF NOT axis1.State.finish OR axis1.State.busy THEN 
		 _updateHmiTextWithAxisBusy(axisName:= axisName1);
	ELSIF NOT axis1.State.pass THEN 
		_addressRestart:= _SubStep.actual;
		_getAxisErrorTexts(name			:= axisName1,
						   description	:= axis1.State.description); 
		_SubStep.set(request:= _SUB_ADDRESS_RETRY_ABORT);
	ELSE 
		_subStep.INC();
	END_IF			
END_IF

(* Home axis Right*)
IF _SubStep.isActive(1) THEN 
	 IF NOT axis2.Ex_Homing() THEN
		 _updateHmiTextWithAxisBusy(axisName:= axisName2);		 
	ELSIF NOT axis2.State.finish OR axis2.State.busy THEN 
		 _updateHmiTextWithAxisBusy(axisName:= axisName2);
	ELSIF NOT axis2.State.pass THEN 
		_addressRestart:= _SubStep.actual;
		_getAxisErrorTexts(name			:= axisName2,
						   description	:= axis2.State.description); 
		_SubStep.set(request:= _SUB_ADDRESS_RETRY_ABORT);
	ELSE 
		_subStep.set(request:= _SUB_ADDRESS_PASS);
	END_IF			
END_IF

(* Pass *)
IF _SubStep.isActive(_SUB_ADDRESS_PASS) THEN 
	_Step.Condition:= TRUE;
END_IF

(* Fail - Retry/Abort *)
IF _SubStep.isActive(_SUB_ADDRESS_RETRY_ABORT) THEN 
	_retryAbort(
		numOfTargetRetries	:= _UNLIMITED_RETRY_NUMBER,
		retryAddress		:= _addressRestart,
		abortAddress		:= _SubStep.actual-1);
END_IF

_step.Control();
END_METHOD

METHOD PROTECTED _a2_X_HomeAxis
VAR_INPUT
	axis			: REFERENCE TO  KOSTAL_AF2024_Drivers_Actuation_Axis_Festo_CMMT_AS.FB_FESTO_CMMT_AS;
	axisName		: KOSTAL_AF2024_Core_Settings.T_MaxString;
END_VAR
IF _step.toggle THEN 
	_stepDescription:= "HomeAxis";
END_IF
(* Is Axis X Home? *) 
IF _SubStep.isActive(0) THEN 
	IF _isHomeDone AND axis.AxisPositionAct = axis.HomingPosition THEN 
		_SubStep.set(request:= _SUB_ADDRESS_PASS);
	ELSE 
		_SubStep.INC();
	END_IF
END_IF
(* Home axis Left*)
IF _SubStep.isActive(1) THEN 
	 IF NOT axis.Ex_Homing() THEN
		 _updateHmiTextWithAxisBusy(axisName:= axisName);		 
	ELSIF NOT axis.State.finish OR axis.State.busy THEN 
		 _updateHmiTextWithAxisBusy(axisName:= axisName);
	ELSIF NOT axis.State.pass THEN 
		_addressRestart:= _SubStep.actual;
		_getAxisErrorTexts(name			:= axisName,
						   description	:= axis.State.description); 
		_SubStep.set(request:= _SUB_ADDRESS_RETRY_ABORT);
	ELSE 
		_SubStep.set(request:= _SUB_ADDRESS_PASS); 
	END_IF			
END_IF

(* Pass *)
IF _SubStep.isActive(_SUB_ADDRESS_PASS) THEN 
	_Step.Condition:= TRUE;
END_IF

(* Fail - Retry/Abort *)
IF _SubStep.isActive(_SUB_ADDRESS_RETRY_ABORT) THEN 
	_retryAbort(
		numOfTargetRetries	:= _UNLIMITED_RETRY_NUMBER,
		retryAddress		:= _addressRestart,
		abortAddress		:= _SubStep.actual-1);
END_IF

_step.Control();
END_METHOD

METHOD PROTECTED _a2_X_HomeAxisTC3
VAR_INPUT
	axis		: I_LinearAxis_position;
	axisName	: KOSTAL_AF2024_Core_Settings.T_MaxString;
END_VAR
IF _step.toggle THEN 
	_stepDescription:= "HomeAxis";
END_IF

//(* Is Axis X Home? *) 
//IF _SubStep.isActive(0) THEN 
//	IF _isHomeDone AND axis.IlinearAxis_PositionAct = axis.IlinearAxis_HomingPosition THEN 
//		_SubStep.set(request:= _SUB_ADDRESS_PASS);
//	ELSE 
//		_SubStep.INC();
//	END_IF
//END_IF

(* Home Axis X *)
 IF _SubStep.isActive(0) THEN 
	 axis.IlinearAxis_Homing();
	 IF NOT axis.IlinearAxis_State.finish THEN 
		 _updateHmiTextWithAxisBusy(axisName:= axisName);
	ELSIF NOT axis.IlinearAxis_State.pass THEN 
		_addressRestart:= _SubStep.actual;
		_getAxisErrorTexts(
			name		:= axisName,
			description	:= STRING_TO_WSTRING(axis.IlinearAxis_State.description));
		_SubStep.set(request:= _SUB_ADDRESS_RETRY_ABORT);
	ELSE 
		_subStep.set(request:= _SUB_ADDRESS_PASS);
	END_IF		
END_IF

(* Pass *)
IF _SubStep.isActive(_SUB_ADDRESS_PASS) THEN 
	_isHomeDone:= TRUE;
	_Step.Condition:= TRUE;
END_IF

(* Fail - Retry/Abort *)
IF _SubStep.isActive(_SUB_ADDRESS_RETRY_ABORT) THEN 
	_retryAbort(
		numOfTargetRetries	:= _UNLIMITED_RETRY_NUMBER,
		retryAddress		:= _addressRestart,
		abortAddress		:= _SubStep.actual-1);
END_IF

_step.Control();
END_METHOD

METHOD PROTECTED _a2_X_InitAxes
VAR_INPUT
	axis1			: REFERENCE TO KOSTAL_AF2024_Drivers_Actuation_Axis_Festo_CMMT_AS.FB_FESTO_CMMT_AS;
	axisName1		: KOSTAL_AF2024_Core_Settings.T_MaxString;
	axis2			: REFERENCE TO KOSTAL_AF2024_Drivers_Actuation_Axis_Festo_CMMT_AS.FB_FESTO_CMMT_AS;
	axisName2		: KOSTAL_AF2024_Core_Settings.T_MaxString;
END_VAR
(* Reset Axis Left *)
IF _SubStep.isActive(0) THEN 
	_addressRestart:= _SubStep.actual;
	IF axis1.Fault THEN 
	axis1.ResetFault();
		IF NOT axis1.AxisError THEN 
			_SubStep.INC();
		ELSE 
			_updateHmiTextWithAxisBusy(axisName:= axisName1); 
		END_IF
	ELSE 
		_SubStep.INC();
	END_IF
END_IF

(* Enable Axis Left *)
IF _SubStep.isActive(1) THEN 
	axis1.Ex_On();
	IF NOT axis1.State.finish THEN 
		_updateHmiTextWithAxisBusy(axisName:= axisName1);
	ELSIF NOT axis1.State.pass THEN 
		_subStepError:= "Left axis in error";
		_subStepMessage:= axis1.State.description;
		_SubStep.set(request:= _SUB_ADDRESS_RETRY_ABORT);
	ELSIF axis1.AxisIsOn THEN 
		_SubStep.INC();
	ELSE 
		_updateHmiTextWithAxisBusy(axisName:= axisName1);
	END_IF
END_IF

